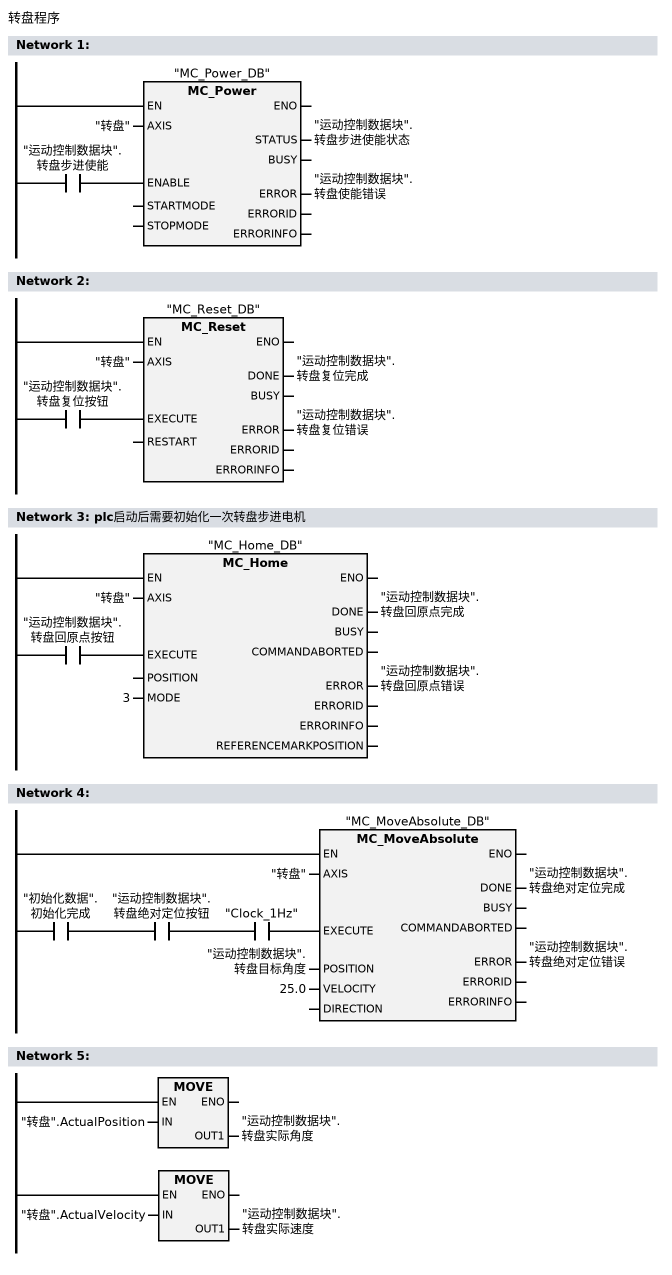
   "MC_Power_DB"(Axis := "转盘",   // MC_Power
                 Enable := "运动控制数据块".转盘步进使能,
                 Status => "运动控制数据块".转盘步进使能状态,
                 Error => "运动控制数据块".转盘使能错误);
END_REGION

REGION Network 2
   "MC_Reset_DB"(Axis := "转盘", Execute := "运动控制数据块".转盘复位按钮, Done => "运动控制数据块".转盘复位完成, Error => "运动控制数据块".转盘复位错误);   // MC_Reset
END_REGION

REGION Network 3: plc启动后需要初始化一次转盘步进电机
   "MC_Home_DB"(Axis := "转盘",   // MC_Home
                Execute := "运动控制数据块".转盘回原点按钮,
                Mode := 3,
                Done => "运动控制数据块".转盘回原点完成,
                Error => "运动控制数据块".转盘回原点错误);
END_REGION

REGION Network 4
   "MC_MoveAbsolute_DB"(Axis := "转盘",   // MC_MoveAbsolute
                        Execute := "初始化数据".初始化完成 AND "运动控制数据块".转盘绝对定位按钮 AND "Clock_1Hz",
                        Position := "运动控制数据块".转盘目标角度,
                        Velocity := 25.0,
                        Done => "运动控制数据块".转盘绝对定位完成,
                        Error => "运动控制数据块".转盘绝对定位错误);
END_REGION

REGION Network 5
   RUNG wire#powerrail
      Move(in := "转盘".ActualPosition, out1 => "运动控制数据块".转盘实际角度)
   END_RUNG
   RUNG wire#powerrail
      Move(in := "转盘".ActualVelocity, out1 => "运动控制数据块".转盘实际速度)
   END_RUNG
   // the same network as SCL:
   "运动控制数据块".转盘实际角度 := "转盘".ActualPosition;
   "运动控制数据块".转盘实际速度 := "转盘".ActualVelocity;
END_REGION
END_FUNCTION

FUNCTION "机械手程序" : Void   // FC8, LAD
{ S7_Optimized_Access := 'TRUE' }
VERSION : 0.1
// 极限位：左100，右-180
BEGIN

REGION Network 1: 轴使能
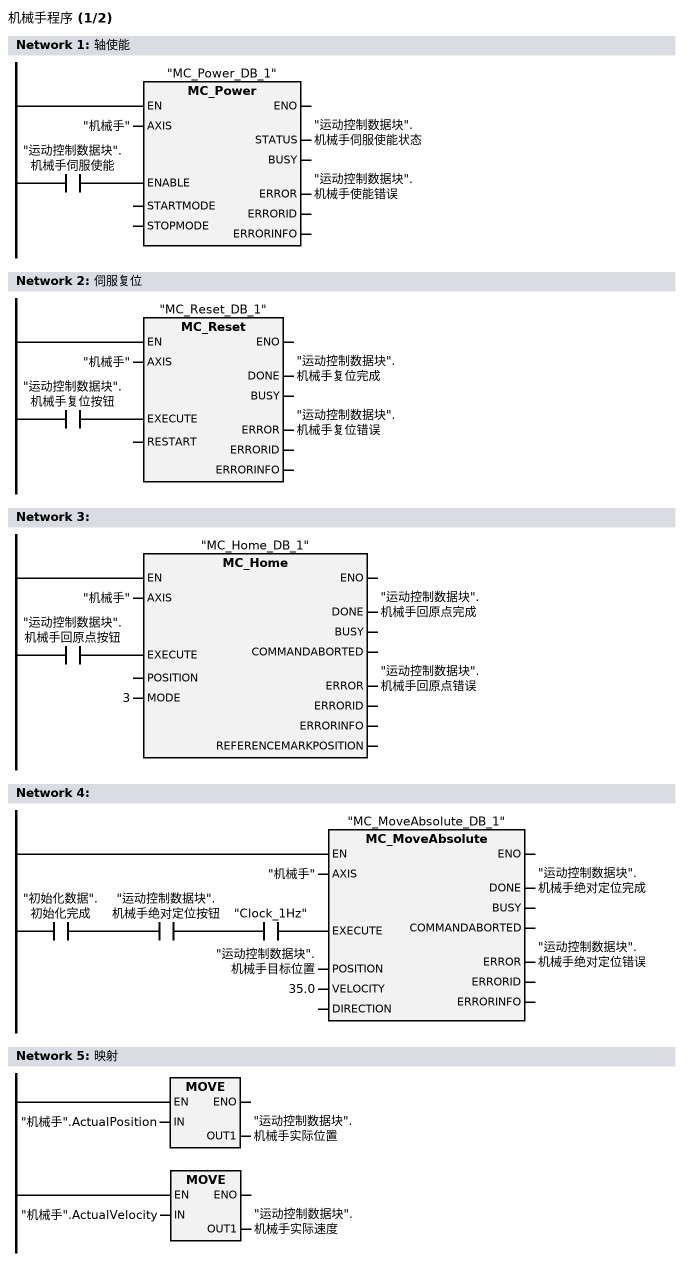
   "MC_Power_DB_1"(Axis := "机械手",   // MC_Power
                   Enable := "运动控制数据块".机械手伺服使能,
                   Status => "运动控制数据块".机械手伺服使能状态,
                   Error => "运动控制数据块".机械手使能错误);
END_REGION

REGION Network 2: 伺服复位
   "MC_Reset_DB_1"(Axis := "机械手",   // MC_Reset
                   Execute := "运动控制数据块".机械手复位按钮,
                   Done => "运动控制数据块".机械手复位完成,
                   Error => "运动控制数据块".机械手复位错误);
END_REGION

REGION Network 3
   "MC_Home_DB_1"(Axis := "机械手",   // MC_Home
                  Execute := "运动控制数据块".机械手回原点按钮,
                  Mode := 3,
                  Done => "运动控制数据块".机械手回原点完成,
                  Error => "运动控制数据块".机械手回原点错误);
END_REGION

REGION Network 4
   "MC_MoveAbsolute_DB_1"(Axis := "机械手",   // MC_MoveAbsolute
                          Execute := "初始化数据".初始化完成 AND "运动控制数据块".机械手绝对定位按钮 AND "Clock_1Hz",
                          Position := "运动控制数据块".机械手目标位置,
                          Velocity := 35.0,
                          Done => "运动控制数据块".机械手绝对定位完成,
                          Error => "运动控制数据块".机械手绝对定位错误);
END_REGION

REGION Network 5: 映射
   RUNG wire#powerrail
      Move(in := "机械手".ActualPosition, out1 => "运动控制数据块".机械手实际位置)
   END_RUNG
   RUNG wire#powerrail
      Move(in := "机械手".ActualVelocity, out1 => "运动控制数据块".机械手实际速度)
   END_RUNG
   // the same network as SCL:
   "运动控制数据块".机械手实际位置 := "机械手".ActualPosition;
   "运动控制数据块".机械手实际速度 := "机械手".ActualVelocity;
END_REGION

REGION Network 6
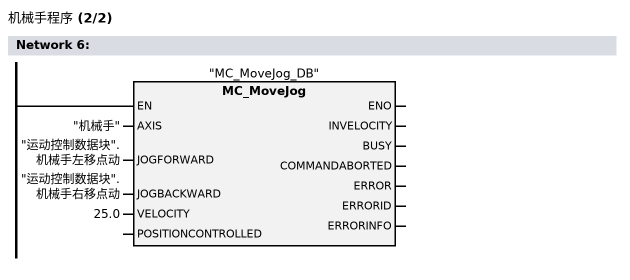
   "MC_MoveJog_DB"(Axis := "机械手",   // MC_MoveJog
                   JogForward := "运动控制数据块".机械手左移点动,
                   JogBackward := "运动控制数据块".机械手右移点动,
                   Velocity := 25.0);
END_REGION
END_FUNCTION

FUNCTION "[00]轴回零" : Void   // FC9, LAD
{ S7_Optimized_Access := 'TRUE' }
VERSION : 0.1
   VAR_TEMP   // added for the SCL form of the ladder/FBD networks
      _w1 : Bool;
   END_VAR
BEGIN

REGION Network 1
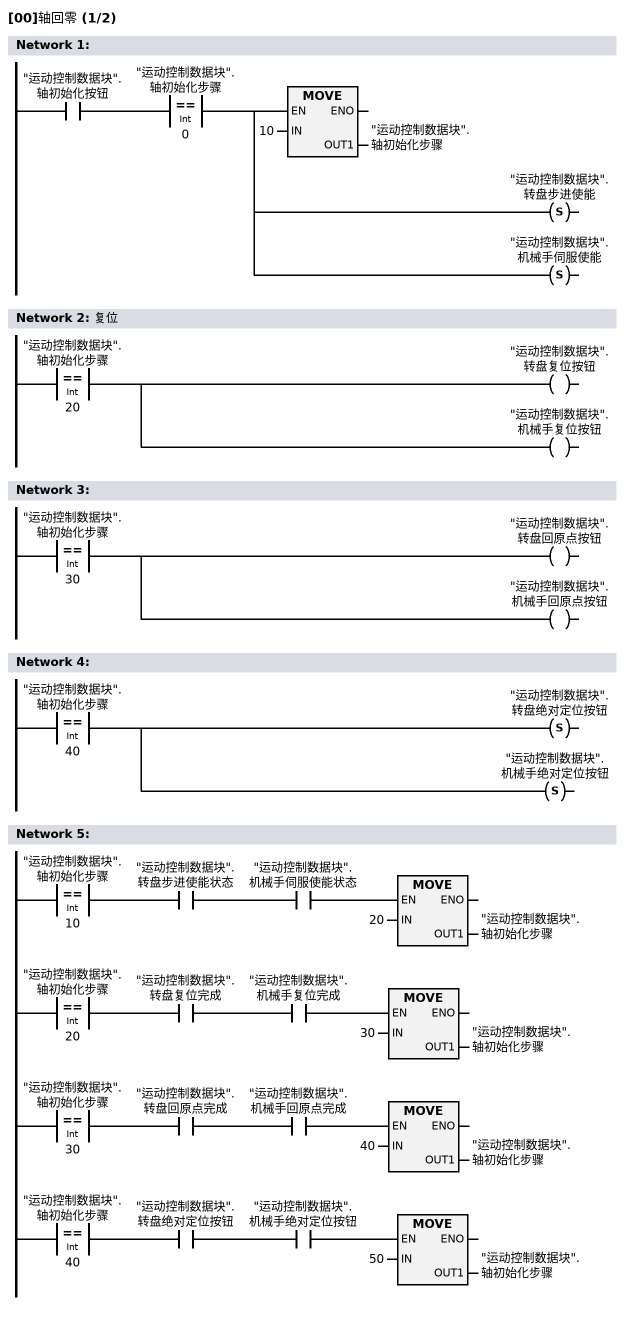
   RUNG wire#powerrail
      Contact( "运动控制数据块".轴初始化按钮 )
      { S7_Templates := "SrcType := Int" } EQ_Contact(in1 := "运动控制数据块".轴初始化步骤, in2 := 0)
      wire#w1
      Move(in := 10, out1 => "运动控制数据块".轴初始化步骤)
   END_RUNG
   RUNG wire#w1
      S_Coil( "运动控制数据块".转盘步进使能 )
   END_RUNG
   RUNG wire#w1
      S_Coil( "运动控制数据块".机械手伺服使能 )
   END_RUNG
   // the same network as SCL:
   #_w1 := "运动控制数据块".轴初始化按钮 AND ("运动控制数据块".轴初始化步骤 = 0);
   IF #_w1 THEN
       "运动控制数据块".轴初始化步骤 := 10;
       "运动控制数据块".转盘步进使能 := TRUE;
       "运动控制数据块".机械手伺服使能 := TRUE;
   END_IF;
END_REGION

REGION Network 2: 复位
   RUNG wire#powerrail
      { S7_Templates := "SrcType := Int" } EQ_Contact(in1 := "运动控制数据块".轴初始化步骤, in2 := 20)
      wire#w1
      Coil( "运动控制数据块".转盘复位按钮 )
   END_RUNG
   RUNG wire#w1
      Coil( "运动控制数据块".机械手复位按钮 )
   END_RUNG
   // the same network as SCL:
   "运动控制数据块".转盘复位按钮 := "运动控制数据块".轴初始化步骤 = 20;
   "运动控制数据块".机械手复位按钮 := "运动控制数据块".转盘复位按钮;
END_REGION

REGION Network 3
   RUNG wire#powerrail
      { S7_Templates := "SrcType := Int" } EQ_Contact(in1 := "运动控制数据块".轴初始化步骤, in2 := 30)
      wire#w1
      Coil( "运动控制数据块".转盘回原点按钮 )
   END_RUNG
   RUNG wire#w1
      Coil( "运动控制数据块".机械手回原点按钮 )
   END_RUNG
   // the same network as SCL:
   "运动控制数据块".转盘回原点按钮 := "运动控制数据块".轴初始化步骤 = 30;
   "运动控制数据块".机械手回原点按钮 := "运动控制数据块".转盘回原点按钮;
END_REGION

REGION Network 4
   RUNG wire#powerrail
      { S7_Templates := "SrcType := Int" } EQ_Contact(in1 := "运动控制数据块".轴初始化步骤, in2 := 40)
      wire#w1
      S_Coil( "运动控制数据块".转盘绝对定位按钮 )
   END_RUNG
   RUNG wire#w1
      S_Coil( "运动控制数据块".机械手绝对定位按钮 )
   END_RUNG
   // the same network as SCL:
   IF "运动控制数据块".轴初始化步骤 = 40 THEN
       "运动控制数据块".转盘绝对定位按钮 := TRUE;
       "运动控制数据块".机械手绝对定位按钮 := TRUE;
   END_IF;
END_REGION

REGION Network 5
   RUNG wire#powerrail
      { S7_Templates := "SrcType := Int" } EQ_Contact(in1 := "运动控制数据块".轴初始化步骤, in2 := 10)
      Contact( "运动控制数据块".转盘步进使能状态 )
      Contact( "运动控制数据块".机械手伺服使能状态 )
      Move(in := 20, out1 => "运动控制数据块".轴初始化步骤)
   END_RUNG
   RUNG wire#powerrail
      { S7_Templates := "SrcType := Int" } EQ_Contact(in1 := "运动控制数据块".轴初始化步骤, in2 := 20)
      Contact( "运动控制数据块".转盘复位完成 )
      Contact( "运动控制数据块".机械手复位完成 )
      Move(in := 30, out1 => "运动控制数据块".轴初始化步骤)
   END_RUNG
   RUNG wire#powerrail
      { S7_Templates := "SrcType := Int" } EQ_Contact(in1 := "运动控制数据块".轴初始化步骤, in2 := 30)
      Contact( "运动控制数据块".转盘回原点完成 )
      Contact( "运动控制数据块".机械手回原点完成 )
      Move(in := 40, out1 => "运动控制数据块".轴初始化步骤)
   END_RUNG
   RUNG wire#powerrail
      { S7_Templates := "SrcType := Int" } EQ_Contact(in1 := "运动控制数据块".轴初始化步骤, in2 := 40)
      Contact( "运动控制数据块".转盘绝对定位按钮 )
      Contact( "运动控制数据块".机械手绝对定位按钮 )
      Move(in := 50, out1 => "运动控制数据块".轴初始化步骤)
   END_RUNG
   // the same network as SCL:
   IF ("运动控制数据块".轴初始化步骤 = 10) AND "运动控制数据块".转盘步进使能状态 AND "运动控制数据块".机械手伺服使能状态 THEN
       "运动控制数据块".轴初始化步骤 := 20;
   END_IF;
   IF ("运动控制数据块".轴初始化步骤 = 20) AND "运动控制数据块".转盘复位完成 AND "运动控制数据块".机械手复位完成 THEN "运动控制数据块".轴初始化步骤 := 30; END_IF;
   IF ("运动控制数据块".轴初始化步骤 = 30) AND "运动控制数据块".转盘回原点完成 AND "运动控制数据块".机械手回原点完成 THEN
       "运动控制数据块".轴初始化步骤 := 40;
   END_IF;
   IF ("运动控制数据块".轴初始化步骤 = 40) AND "运动控制数据块".转盘绝对定位按钮 AND "运动控制数据块".机械手绝对定位按钮 THEN
       "运动控制数据块".轴初始化步骤 := 50;
   END_IF;
END_REGION

REGION Network 6: 轴初始化完成
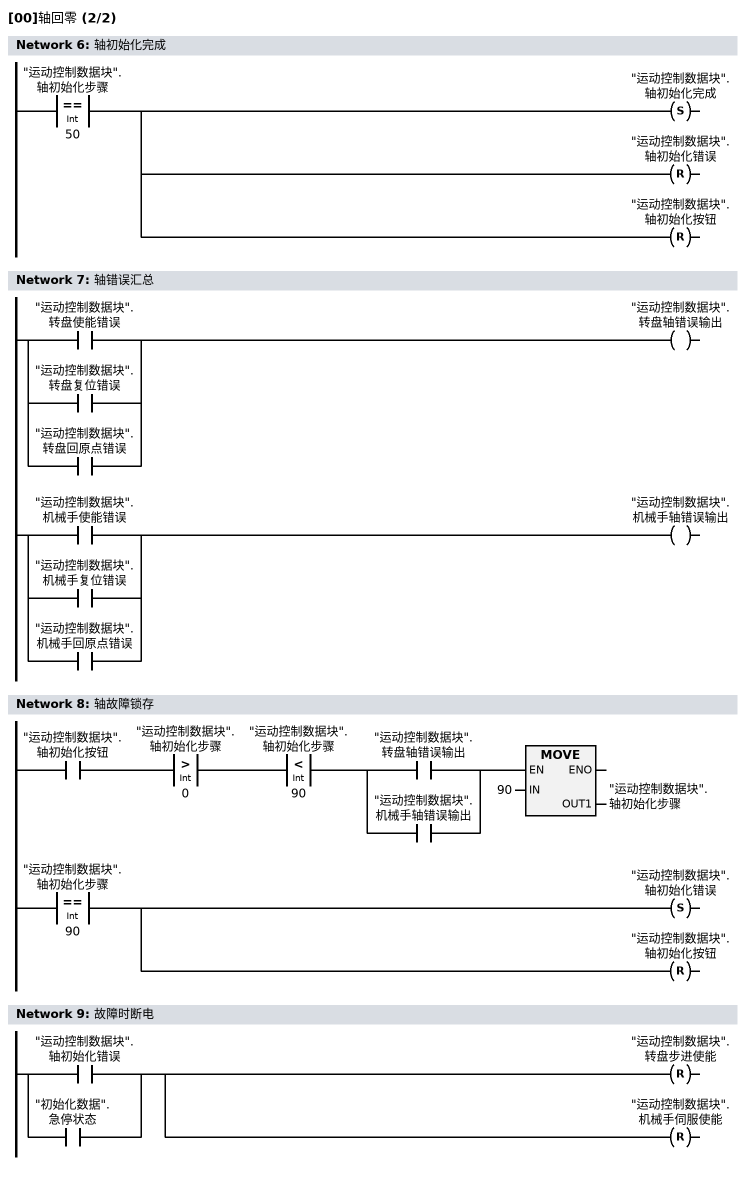
   RUNG wire#powerrail
      { S7_Templates := "SrcType := Int" } EQ_Contact(in1 := "运动控制数据块".轴初始化步骤, in2 := 50)
      wire#w1
      S_Coil( "运动控制数据块".轴初始化完成 )
   END_RUNG
   RUNG wire#w1
      R_Coil( "运动控制数据块".轴初始化错误 )
   END_RUNG
   RUNG wire#w1
      R_Coil( "运动控制数据块".轴初始化按钮 )
   END_RUNG
   // the same network as SCL:
   IF "运动控制数据块".轴初始化步骤 = 50 THEN
       "运动控制数据块".轴初始化完成 := TRUE;
       "运动控制数据块".轴初始化错误 := FALSE;
       "运动控制数据块".轴初始化按钮 := FALSE;
   END_IF;
END_REGION

REGION Network 7: 轴错误汇总
   RUNG wire#powerrail
      Contact( "运动控制数据块".转盘使能错误 )
      wire#w1
      Coil( "运动控制数据块".转盘轴错误输出 )
   END_RUNG
   RUNG wire#powerrail
      Contact( "运动控制数据块".转盘复位错误 )
   END_RUNG wire#w1
   RUNG wire#powerrail
      Contact( "运动控制数据块".转盘回原点错误 )
   END_RUNG wire#w1
   RUNG wire#powerrail
      Contact( "运动控制数据块".机械手使能错误 )
      wire#w2
      Coil( "运动控制数据块".机械手轴错误输出 )
   END_RUNG
   RUNG wire#powerrail
      Contact( "运动控制数据块".机械手复位错误 )
   END_RUNG wire#w2
   RUNG wire#powerrail
      Contact( "运动控制数据块".机械手回原点错误 )
   END_RUNG wire#w2
   // the same network as SCL:
   "运动控制数据块".转盘轴错误输出 := "运动控制数据块".转盘使能错误 OR "运动控制数据块".转盘复位错误 OR "运动控制数据块".转盘回原点错误;
   "运动控制数据块".机械手轴错误输出 := "运动控制数据块".机械手使能错误 OR "运动控制数据块".机械手复位错误 OR "运动控制数据块".机械手回原点错误;
END_REGION

REGION Network 8: 轴故障锁存
   RUNG wire#powerrail
      Contact( "运动控制数据块".轴初始化按钮 )
      { S7_Templates := "SrcType := Int" } GT_Contact(in1 := "运动控制数据块".轴初始化步骤, in2 := 0)
      { S7_Templates := "SrcType := Int" } LT_Contact(in1 := "运动控制数据块".轴初始化步骤, in2 := 90)
      wire#w1
      Contact( "运动控制数据块".转盘轴错误输出 )
      wire#w2
      Move(in := 90, out1 => "运动控制数据块".轴初始化步骤)
   END_RUNG
   RUNG wire#w1
      Contact( "运动控制数据块".机械手轴错误输出 )
   END_RUNG wire#w2
   RUNG wire#powerrail
      { S7_Templates := "SrcType := Int" } EQ_Contact(in1 := "运动控制数据块".轴初始化步骤, in2 := 90)
      wire#w3
      S_Coil( "运动控制数据块".轴初始化错误 )
   END_RUNG
   RUNG wire#w3
      R_Coil( "运动控制数据块".轴初始化按钮 )
   END_RUNG
   // the same network as SCL:
   IF "运动控制数据块".轴初始化按钮 AND ("运动控制数据块".轴初始化步骤 > 0) AND ("运动控制数据块".轴初始化步骤 < 90) AND ("运动控制数据块".转盘轴错误输出 OR "运动控制数据块".机械手轴错误输出) THEN
       "运动控制数据块".轴初始化步骤 := 90;
   END_IF;
   IF "运动控制数据块".轴初始化步骤 = 90 THEN
       "运动控制数据块".轴初始化错误 := TRUE;
       "运动控制数据块".轴初始化按钮 := FALSE;
   END_IF;
END_REGION

REGION Network 9: 故障时断电
   RUNG wire#powerrail
      Contact( "运动控制数据块".轴初始化错误 )
      wire#w1
      R_Coil( "运动控制数据块".转盘步进使能 )
   END_RUNG
   RUNG wire#powerrail
      Contact( "初始化数据".急停状态 )
   END_RUNG wire#w1
   RUNG wire#w1
      R_Coil( "运动控制数据块".机械手伺服使能 )
   END_RUNG
   // the same network as SCL:
   IF "运动控制数据块".轴初始化错误 OR "初始化数据".急停状态 THEN
       "运动控制数据块".转盘步进使能 := FALSE;
       "运动控制数据块".机械手伺服使能 := FALSE;
   END_IF;
END_REGION
END_FUNCTION

// folder: 通讯数据

FUNCTION "产线通讯" : Void   // FC16, LAD
{ S7_Optimized_Access := 'TRUE' }
VERSION : 0.1
BEGIN

REGION Network 1: 心跳
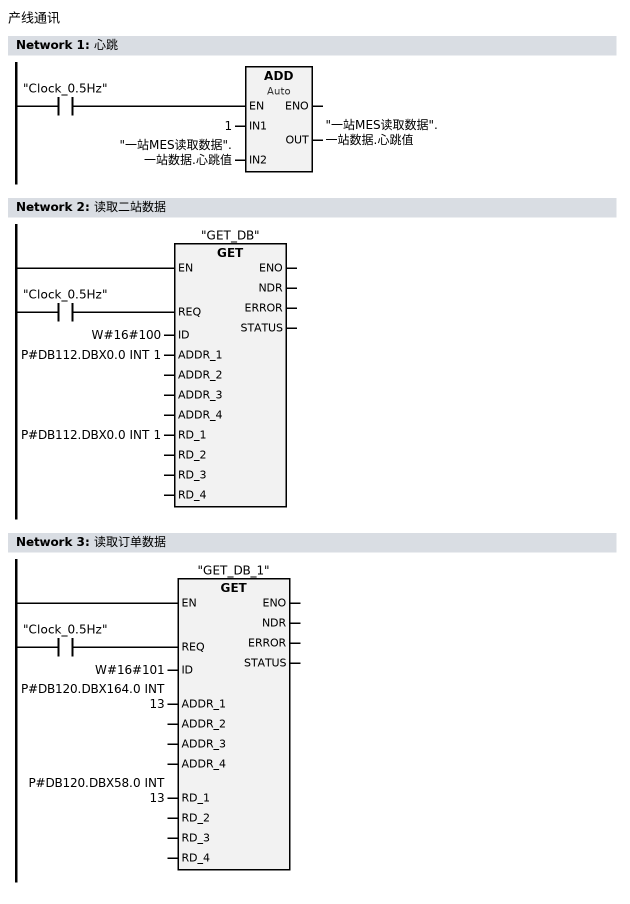
   RUNG wire#powerrail
      Contact( "Clock_0.5Hz" )
      Add(in1 := 1, in2 := "一站MES读取数据".一站数据.心跳值, out => "一站MES读取数据".一站数据.心跳值)
   END_RUNG
   // the same network as SCL:
   IF "Clock_0.5Hz" THEN "一站MES读取数据".一站数据.心跳值 := 1 + "一站MES读取数据".一站数据.心跳值; END_IF;
END_REGION

REGION Network 2: 读取二站数据
   "GET_DB"(REQ := "Clock_0.5Hz", ID := W#16#100, ADDR_1 := P#DB112.DBX0.0 INT 1, RD_1 := P#DB112.DBX0.0 INT 1);   // GET
END_REGION

REGION Network 3: 读取订单数据
   "GET_DB_1"(REQ := "Clock_0.5Hz",   // GET
              ID := W#16#101,
              ADDR_1 := P#DB120.DBX164.0 INT 13,
              RD_1 := P#DB120.DBX58.0 INT 13);
END_REGION
END_FUNCTION

FUNCTION "MES数据映射" : Void   // FC18, LAD
{ S7_Optimized_Access := 'TRUE' }
VERSION : 0.1
BEGIN

REGION Network 1: 运行模式
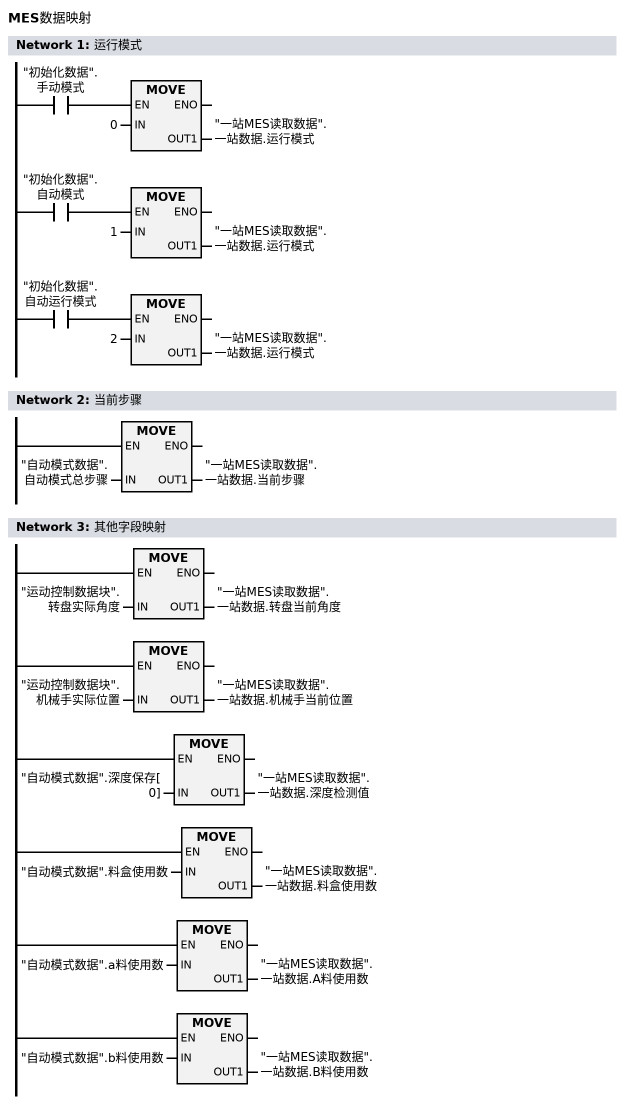
   RUNG wire#powerrail
      Contact( "初始化数据".手动模式 )
      Move(in := 0, out1 => "一站MES读取数据".一站数据.运行模式)
   END_RUNG
   RUNG wire#powerrail
      Contact( "初始化数据".自动模式 )
      Move(in := 1, out1 => "一站MES读取数据".一站数据.运行模式)
   END_RUNG
   RUNG wire#powerrail
      Contact( "初始化数据".自动运行模式 )
      Move(in := 2, out1 => "一站MES读取数据".一站数据.运行模式)
   END_RUNG
   // the same network as SCL:
   IF "初始化数据".手动模式 THEN "一站MES读取数据".一站数据.运行模式 := 0; END_IF;
   IF "初始化数据".自动模式 THEN "一站MES读取数据".一站数据.运行模式 := 1; END_IF;
   IF "初始化数据".自动运行模式 THEN "一站MES读取数据".一站数据.运行模式 := 2; END_IF;
END_REGION

REGION Network 2: 当前步骤
   RUNG wire#powerrail
      Move(in := "自动模式数据".自动模式总步骤, out1 => "一站MES读取数据".一站数据.当前步骤)
   END_RUNG
   // the same network as SCL:
   "一站MES读取数据".一站数据.当前步骤 := "自动模式数据".自动模式总步骤;
END_REGION

REGION Network 3: 其他字段映射
   RUNG wire#powerrail
      Move(in := "运动控制数据块".转盘实际角度, out1 => "一站MES读取数据".一站数据.转盘当前角度)
   END_RUNG
   RUNG wire#powerrail
      Move(in := "运动控制数据块".机械手实际位置, out1 => "一站MES读取数据".一站数据.机械手当前位置)
   END_RUNG
   RUNG wire#powerrail
      Move(in := "自动模式数据".深度保存[0], out1 => "一站MES读取数据".一站数据.深度检测值)
   END_RUNG
   RUNG wire#powerrail
      Move(in := "自动模式数据".料盒使用数, out1 => "一站MES读取数据".一站数据.料盒使用数)
   END_RUNG
   RUNG wire#powerrail
      Move(in := "自动模式数据".a料使用数, out1 => "一站MES读取数据".一站数据.A料使用数)
   END_RUNG
   RUNG wire#powerrail
      Move(in := "自动模式数据".b料使用数, out1 => "一站MES读取数据".一站数据.B料使用数)
   END_RUNG
   // the same network as SCL:
   "一站MES读取数据".一站数据.转盘当前角度 := "运动控制数据块".转盘实际角度;
   "一站MES读取数据".一站数据.机械手当前位置 := "运动控制数据块".机械手实际位置;
   "一站MES读取数据".一站数据.深度检测值 := "自动模式数据".深度保存[0];
   "一站MES读取数据".一站数据.料盒使用数 := "自动模式数据".料盒使用数;
   "一站MES读取数据".一站数据.A料使用数 := "自动模式数据".a料使用数;
   "一站MES读取数据".一站数据.B料使用数 := "自动模式数据".b料使用数;
END_REGION
END_FUNCTION

FUNCTION "扫码器通信" : Void   // FC19, LAD
{ S7_Optimized_Access := 'TRUE' }
VERSION : 0.1
BEGIN

REGION Network 1
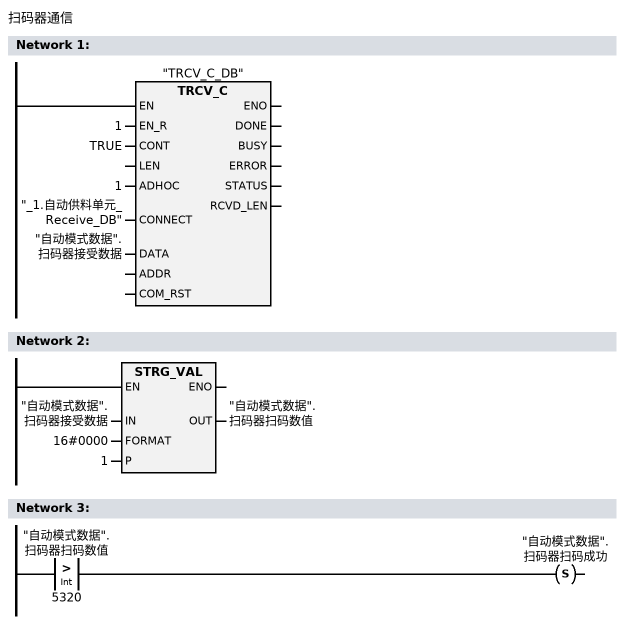
   "TRCV_C_DB"(EN_R := 1, CONT := TRUE, ADHOC := 1, CONNECT := "_1.自动供料单元_Receive_DB", DATA := "自动模式数据".扫码器接受数据);   // TRCV_C
END_REGION

REGION Network 2
   STRG_VAL(IN := "自动模式数据".扫码器接受数据, FORMAT := 16#0000, P := 1, OUT => "自动模式数据".扫码器扫码数值);
END_REGION

REGION Network 3
   RUNG wire#powerrail
      { S7_Templates := "SrcType := Int" } GT_Contact(in1 := "自动模式数据".扫码器扫码数值, in2 := 5320)
      S_Coil( "自动模式数据".扫码器扫码成功 )
   END_RUNG
   // the same network as SCL:
   IF "自动模式数据".扫码器扫码数值 > 5320 THEN "自动模式数据".扫码器扫码成功 := TRUE; END_IF;
END_REGION
END_FUNCTION

FUNCTION "虚实联动映射" : Void   // FC20, LAD
{ S7_Optimized_Access := 'TRUE' }
VERSION : 0.1
BEGIN

REGION Network 1
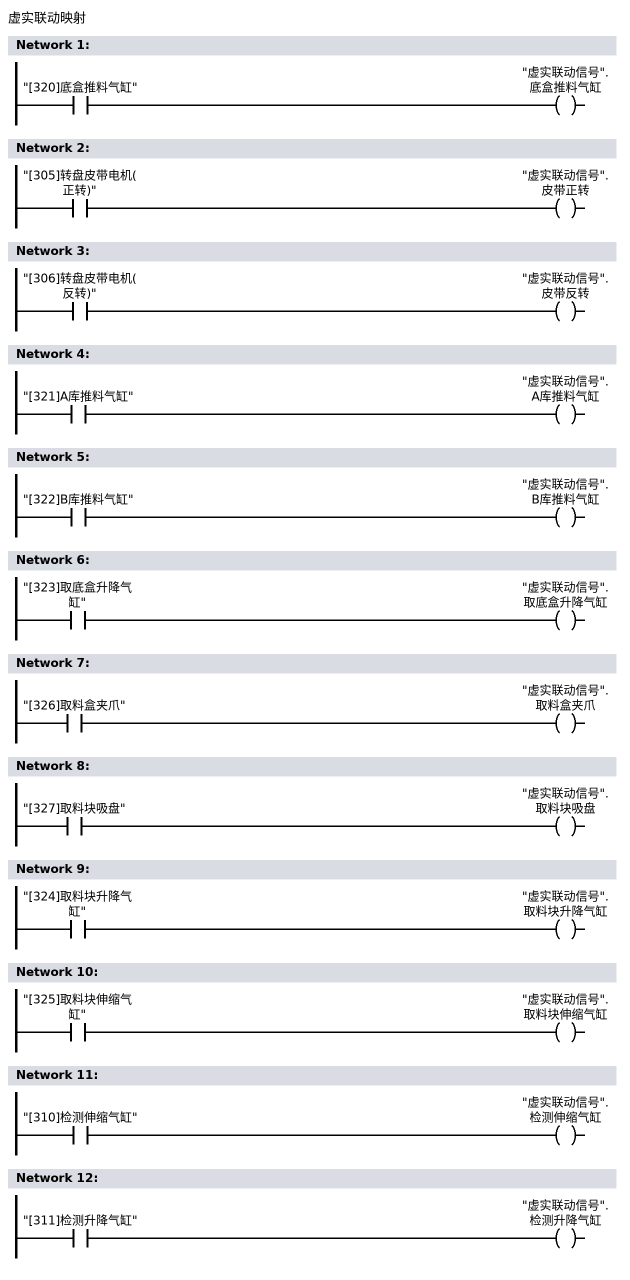
   RUNG wire#powerrail
      Contact( "[320]底盒推料气缸" )
      Coil( "虚实联动信号".底盒推料气缸 )
   END_RUNG
   // the same network as SCL:
   "虚实联动信号".底盒推料气缸 := "[320]底盒推料气缸";
END_REGION

REGION Network 2
   RUNG wire#powerrail
      Contact( "[305]转盘皮带电机(正转)" )
      Coil( "虚实联动信号".皮带正转 )
   END_RUNG
   // the same network as SCL:
   "虚实联动信号".皮带正转 := "[305]转盘皮带电机(正转)";
END_REGION

REGION Network 3
   RUNG wire#powerrail
      Contact( "[306]转盘皮带电机(反转)" )
      Coil( "虚实联动信号".皮带反转 )
   END_RUNG
   // the same network as SCL:
   "虚实联动信号".皮带反转 := "[306]转盘皮带电机(反转)";
END_REGION

REGION Network 4
   RUNG wire#powerrail
      Contact( "[321]A库推料气缸" )
      Coil( "虚实联动信号".A库推料气缸 )
   END_RUNG
   // the same network as SCL:
   "虚实联动信号".A库推料气缸 := "[321]A库推料气缸";
END_REGION

REGION Network 5
   RUNG wire#powerrail
      Contact( "[322]B库推料气缸" )
      Coil( "虚实联动信号".B库推料气缸 )
   END_RUNG
   // the same network as SCL:
   "虚实联动信号".B库推料气缸 := "[322]B库推料气缸";
END_REGION

REGION Network 6
   RUNG wire#powerrail
      Contact( "[323]取底盒升降气缸" )
      Coil( "虚实联动信号".取底盒升降气缸 )
   END_RUNG
   // the same network as SCL:
   "虚实联动信号".取底盒升降气缸 := "[323]取底盒升降气缸";
END_REGION

REGION Network 7
   RUNG wire#powerrail
      Contact( "[326]取料盒夹爪" )
      Coil( "虚实联动信号".取料盒夹爪 )
   END_RUNG
   // the same network as SCL:
   "虚实联动信号".取料盒夹爪 := "[326]取料盒夹爪";
END_REGION

REGION Network 8
   RUNG wire#powerrail
      Contact( "[327]取料块吸盘" )
      Coil( "虚实联动信号".取料块吸盘 )
   END_RUNG
   // the same network as SCL:
   "虚实联动信号".取料块吸盘 := "[327]取料块吸盘";
END_REGION

REGION Network 9
   RUNG wire#powerrail
      Contact( "[324]取料块升降气缸" )
      Coil( "虚实联动信号".取料块升降气缸 )
   END_RUNG
   // the same network as SCL:
   "虚实联动信号".取料块升降气缸 := "[324]取料块升降气缸";
END_REGION

REGION Network 10
   RUNG wire#powerrail
      Contact( "[325]取料块伸缩气缸" )
      Coil( "虚实联动信号".取料块伸缩气缸 )
   END_RUNG
   // the same network as SCL:
   "虚实联动信号".取料块伸缩气缸 := "[325]取料块伸缩气缸";
END_REGION

REGION Network 11
   RUNG wire#powerrail
      Contact( "[310]检测伸缩气缸" )
      Coil( "虚实联动信号".检测伸缩气缸 )
   END_RUNG
   // the same network as SCL:
   "虚实联动信号".检测伸缩气缸 := "[310]检测伸缩气缸";
END_REGION

REGION Network 12
   RUNG wire#powerrail
      Contact( "[311]检测升降气缸" )
      Coil( "虚实联动信号".检测升降气缸 )
   END_RUNG
   // the same network as SCL:
   "虚实联动信号".检测升降气缸 := "[311]检测升降气缸";
END_REGION
END_FUNCTION

// ===== PLC "2.智能分拣单元"  CPU 1214C DC/DC/DC =====

VAR_GLOBAL   // PLC tag table "默认变量表"
   "System_Byte" AT %MB501 : Byte;
   "FirstScan" AT %M501.0 : Bool;
   "DiagStatusUpdate" AT %M501.1 : Bool;
   "AlwaysTRUE" AT %M501.2 : Bool;
   "AlwaysFALSE" AT %M501.3 : Bool;
   "Clock_Byte" AT %MB500 : Byte;
   "Clock_10Hz" AT %M500.0 : Bool;
   "Clock_5Hz" AT %M500.1 : Bool;
   "Clock_2.5Hz" AT %M500.2 : Bool;
   "Clock_2Hz" AT %M500.3 : Bool;
   "Clock_1.25Hz" AT %M500.4 : Bool;
   "Clock_1Hz" AT %M500.5 : Bool;
   "Clock_0.625Hz" AT %M500.6 : Bool;
   "Clock_0.5Hz" AT %M500.7 : Bool;
   "Tag_1" AT %M5.1 : Bool;
   "注释按钮" AT %M100.0 : Bool;
END_VAR

VAR_GLOBAL   // PLC tag table "第二站变量表"
   "[100]启动" AT %I0.0 : Bool;
   "[101]停止" AT %I0.1 : Bool;
   "[102]复位" AT %I0.2 : Bool;
   "[103]急停" AT %I0.3 : Bool;
   "[104]手自动" AT %I0.4 : Bool;
   "[105]8mm钢球检测" AT %I0.5 : Bool;
   "[107]备用" AT %I0.7 : Bool;
   "[110]备用" AT %I1.0 : Bool;
   "[111]备用" AT %I1.1 : Bool;
   "[112]备用" AT %I1.2 : Bool;
   "[113]备用" AT %I1.3 : Bool;
   "[114]备用" AT %I1.4 : Bool;
   "[120]8mm挡停缩回" AT %I2.0 : Bool;
   "[121]8mm挡停伸出" AT %I2.1 : Bool;
   "[122]8mm料盒到达" AT %I2.2 : Bool;
   "[123]8mm推料缩回" AT %I2.3 : Bool;
   "传输伺服_Drive_OUT" AT %Q64.0 : "PD_TEL3_OUT";
   "[300]8mm分拣步进_脉冲" AT %Q0.0 : Bool;
   "[301]10mm分拣步进_脉冲" AT %Q0.1 : Bool;
   "[302]8mm分拣步进_方向" AT %Q0.2 : Bool;
   "[303]10mm分拣步进_方向" AT %Q0.3 : Bool;
   "[320]8mm挡停气缸" AT %Q2.0 : Bool;
   "[321]8mm推料气缸" AT %Q2.1 : Bool;   // 0为伸出，1为缩回，伸出时料仓检测有效
   "[322]10mm挡停气缸" AT %Q2.2 : Bool;
   "[323]10mm推料气缸" AT %Q2.3 : Bool;
   "[324]备用" AT %Q2.4 : Bool;
   "[325]备用" AT %Q2.5 : Bool;
   "[326]备用" AT %Q2.6 : Bool;
   "[327]备用" AT %Q2.7 : Bool;
   "[124]8mm柱状料仓有无" AT %I2.4 : Bool;
   "[125]10mm挡停缩回" AT %I2.5 : Bool;
   "[115]备用" AT %I1.5 : Bool;
   "[106]10mm钢球检测" AT %I0.6 : Bool;
   "[304]黄色指示灯" AT %Q0.4 : Bool;
   "[305]绿色指示灯" AT %Q0.5 : Bool;
   "[306]红色指示灯" AT %Q0.6 : Bool;
   "[307]声光报警" AT %Q0.7 : Bool;
   "[310]备用" AT %Q1.0 : Bool;
   "[311]备用" AT %Q1.1 : Bool;
   "[156]光栅开关" AT %I5.6 : Bool;
   "[164]深度检测" AT %IW64 : Word;
   "传输伺服_Drive_IN(1)" AT %I68.0 : "PD_TEL3_IN";
   "[126]10mm挡停伸出" AT %I2.6 : Bool;
   "[127]10mm料盒到达" AT %I2.7 : Bool;
   "[130]10mm推料缩回" AT %I3.0 : Bool;
   "[131]10mm柱状料仓有无" AT %I3.1 : Bool;
END_VAR

DATA_BLOCK "初始化数据"   // DB19
{ S7_Optimized_Access := 'FALSE' }
VERSION : 0.1
   VAR
      初始化步骤 : Int;
      初始化完成 : Bool;
      初始化中 : Bool;
      初始化故障 : Bool;
      急停状态 : Bool;
      复位完成 : Bool;
      手动模式 : Bool;
      自动模式 : Bool;
      自动运行模式 : Bool;
      黄灯_内部 : Bool;
      红灯_内部 : Bool;
      绿灯_内部 : Bool;
      安全光栅被挡 : Bool;
      报警等级 : Int;
      报警确认按钮 : Bool;
      "8mm挡停气缸报警" : Bool;
      "10mm挡停气缸报警" : Bool;
      报警总输出 : Bool;
      报警状态确认 : Bool;
   END_VAR
BEGIN
END_DATA_BLOCK

DATA_BLOCK "状态控制数据"   // DB28
{ S7_Optimized_Access := 'FALSE' }
VERSION : 0.1
   VAR
      在线状态 : Bool;
      空闲状态 : Bool;
      忙碌状态 : Bool;
      故障状态 : Bool;
   END_VAR
BEGIN
END_DATA_BLOCK

DATA_BLOCK "二站MES读取数据"   // DB120
{ S7_Optimized_Access := 'FALSE' }
VERSION : 0.1
   VAR
      二站数据 : Struct
         在线状态 : Int;
         运行模式 : Int;   // 0 手动 / 1 自动待机 / 2 自动运行
         忙碌状态 : Int;   // 0 空闲 / 1 忙碌
         故障状态 : Int;   // 0 = 无故障
         当前订单ID : Int;   // 当前处理的订单
         当前步骤 : Real;
         心跳值 : Int;
         二站完成 : Bool;
         保留 : Bool;
         保留_1 : Bool;
         保留_2 : Bool;
         保留_3 : Bool;
         保留_4 : Bool;
         保留_5 : Bool;
         保留_6 : Bool;
         二站扫码数据 : Int;
         "8mm已灌注数量" : Int;
         "10mm已灌注数量" : Int;
         "8mml料仓钢珠有无" : Bool;   // 1有0无
         "10mm料仓钢珠有无" : Bool;   // 1有0无
         二站保留数据 : Array[0..9] of Int;
      END_STRUCT;
      订单数据 : Struct
         订单id : Int;
         ab物料 : Int;   // 1A，2B，3不需要
         小钢珠数量 : Int;
         大钢珠数量 : Int;
         存储仓位 : Int;
         当前订单完成 : Bool;
         开始信号 : Int;
         复位信号 : Int;
         订单保留数据 : Array[0..4] of Int;
      END_STRUCT;
   END_VAR
BEGIN
END_DATA_BLOCK

// folder: System blocks/Program resources

DATA_BLOCK "IEC_Timer_0_DB_16"   // DB3
{ S7_Optimized_Access := 'TRUE' }
AUTHOR : Simatic
FAMILY : IEC
NAME : IEC_TMR
VERSION : 1.0
// stored: InstanceOfName IEC_TIMER
"IEC_TIMER"
BEGIN
END_DATA_BLOCK

DATA_BLOCK "IEC_Timer_0_DB"   // DB4
{ S7_Optimized_Access := 'TRUE' }
AUTHOR : Simatic
FAMILY : IEC
NAME : IEC_TMR
VERSION : 1.0
// stored: InstanceOfName IEC_TIMER
"IEC_TIMER"
BEGIN
END_DATA_BLOCK

DATA_BLOCK "IEC_Timer_0_DB_1"   // DB5
{ S7_Optimized_Access := 'TRUE' }
AUTHOR : Simatic
FAMILY : IEC
NAME : IEC_TMR
VERSION : 1.0
// stored: InstanceOfName IEC_TIMER
"IEC_TIMER"
BEGIN
END_DATA_BLOCK

DATA_BLOCK "IEC_Timer_0_DB_2"   // DB7
{ S7_Optimized_Access := 'TRUE' }
AUTHOR : Simatic
FAMILY : IEC
NAME : IEC_TMR
VERSION : 1.0
// stored: InstanceOfName IEC_TIMER
"IEC_TIMER"
BEGIN
END_DATA_BLOCK

DATA_BLOCK "IEC_Timer_0_DB_3"   // DB8
{ S7_Optimized_Access := 'TRUE' }
AUTHOR : Simatic
FAMILY : IEC
NAME : IEC_TMR
VERSION : 1.0
// stored: InstanceOfName IEC_TIMER
"IEC_TIMER"
BEGIN
END_DATA_BLOCK

DATA_BLOCK "IEC_Timer_0_DB_4"   // DB9
{ S7_Optimized_Access := 'TRUE' }
AUTHOR : Simatic
FAMILY : IEC
NAME : IEC_TMR
VERSION : 1.0
// stored: InstanceOfName IEC_TIMER
"IEC_TIMER"
BEGIN
END_DATA_BLOCK

DATA_BLOCK "IEC_Timer_0_DB_5"   // DB10
{ S7_Optimized_Access := 'TRUE' }
AUTHOR : Simatic
FAMILY : IEC
NAME : IEC_TMR
VERSION : 1.0
// stored: InstanceOfName IEC_TIMER
"IEC_TIMER"
BEGIN
END_DATA_BLOCK

DATA_BLOCK "IEC_Timer_0_DB_6"   // DB11
{ S7_Optimized_Access := 'TRUE' }
AUTHOR : Simatic
FAMILY : IEC
NAME : IEC_TMR
VERSION : 1.0
// stored: InstanceOfName IEC_TIMER
"IEC_TIMER"
BEGIN
END_DATA_BLOCK

DATA_BLOCK "IEC_Timer_0_DB_7"   // DB12
{ S7_Optimized_Access := 'TRUE' }
AUTHOR : Simatic
FAMILY : IEC
NAME : IEC_TMR
VERSION : 1.0
// stored: InstanceOfName IEC_TIMER
"IEC_TIMER"
BEGIN
END_DATA_BLOCK

DATA_BLOCK "IEC_Timer_0_DB_8"   // DB13
{ S7_Optimized_Access := 'TRUE' }
AUTHOR : Simatic
FAMILY : IEC
NAME : IEC_TMR
VERSION : 1.0
// stored: InstanceOfName IEC_TIMER
"IEC_TIMER"
BEGIN
END_DATA_BLOCK

DATA_BLOCK "IEC_Timer_0_DB_9"   // DB14
{ S7_Optimized_Access := 'TRUE' }
AUTHOR : Simatic
FAMILY : IEC
NAME : IEC_TMR
VERSION : 1.0
// stored: InstanceOfName IEC_TIMER
"IEC_TIMER"
BEGIN
END_DATA_BLOCK

DATA_BLOCK "_2.智能分拣单元_Receive_DB"   // DB16
{ S7_Optimized_Access := 'TRUE' }
AUTHOR : SIMATIC
FAMILY : MC7Plus
NAME : TC_IP_v4
VERSION : 1.0
// stored: InstanceOfName TCON_IP_v4
"TCON_IP_v4"
BEGIN
   ID := 110;
   InterfaceId := 64;
   LocalPort := 8899;
   RemotePort := 8899;
   RemoteAddress.ADDR[1] := 192;
   RemoteAddress.ADDR[2] := 168;
   RemoteAddress.ADDR[3] := 40;
   RemoteAddress.ADDR[4] := 101;
END_DATA_BLOCK

DATA_BLOCK "IEC_Timer_0_DB_10"   // DB17
{ S7_Optimized_Access := 'TRUE' }
AUTHOR : Simatic
FAMILY : IEC
NAME : IEC_TMR
VERSION : 1.0
// stored: InstanceOfName IEC_TIMER
"IEC_TIMER"
BEGIN
END_DATA_BLOCK

DATA_BLOCK "IEC_Timer_0_DB_11"   // DB18
{ S7_Optimized_Access := 'TRUE' }
AUTHOR : Simatic
FAMILY : IEC
NAME : IEC_TMR
VERSION : 1.0
// stored: InstanceOfName IEC_TIMER
"IEC_TIMER"
BEGIN
END_DATA_BLOCK

DATA_BLOCK "IEC_Timer_0_DB_12"   // DB20
{ S7_Optimized_Access := 'TRUE' }
AUTHOR : Simatic
FAMILY : IEC
NAME : IEC_TMR
VERSION : 1.0
// stored: InstanceOfName IEC_TIMER
"IEC_TIMER"
BEGIN
END_DATA_BLOCK

DATA_BLOCK "IEC_Timer_0_DB_13"   // DB21
{ S7_Optimized_Access := 'TRUE' }
AUTHOR : Simatic
FAMILY : IEC
NAME : IEC_TMR
VERSION : 1.0
// stored: InstanceOfName IEC_TIMER
"IEC_TIMER"
BEGIN
END_DATA_BLOCK

DATA_BLOCK "IEC_Timer_0_DB_14"   // DB22
{ S7_Optimized_Access := 'TRUE' }
AUTHOR : Simatic
FAMILY : IEC
NAME : IEC_TMR
VERSION : 1.0
// stored: InstanceOfName IEC_TIMER
"IEC_TIMER"
BEGIN
END_DATA_BLOCK

DATA_BLOCK "IEC_Timer_0_DB_15"   // DB23
{ S7_Optimized_Access := 'TRUE' }
AUTHOR : Simatic
FAMILY : IEC
NAME : IEC_TMR
VERSION : 1.0
// stored: InstanceOfName IEC_TIMER
"IEC_TIMER"
BEGIN
END_DATA_BLOCK

DATA_BLOCK "IEC_Timer_0_DB_19"   // DB25
{ S7_Optimized_Access := 'TRUE' }
AUTHOR : Simatic
FAMILY : IEC
NAME : IEC_TMR
VERSION : 1.0
// stored: InstanceOfName IEC_TIMER
"IEC_TIMER"
BEGIN
END_DATA_BLOCK

DATA_BLOCK "IEC_Timer_0_DB_17"   // DB26
{ S7_Optimized_Access := 'TRUE' }
AUTHOR : Simatic
FAMILY : IEC
NAME : IEC_TMR
VERSION : 1.0
// stored: InstanceOfName IEC_TIMER
"IEC_TIMER"
BEGIN
END_DATA_BLOCK

DATA_BLOCK "IEC_Timer_0_DB_18"   // DB27
{ S7_Optimized_Access := 'TRUE' }
AUTHOR : Simatic
FAMILY : IEC
NAME : IEC_TMR
VERSION : 1.0
// stored: InstanceOfName IEC_TIMER
"IEC_TIMER"
BEGIN
END_DATA_BLOCK

// folder: 手动模式

DATA_BLOCK "手动模式数据"   // DB1
{ S7_Optimized_Access := 'FALSE' }
VERSION : 0.1
   VAR
      手动灌注总步骤 : Real;
      "8mm灌料步骤" : Real;
      "8mm现有钢珠" : Int;
      "8mm目标数量" : Int;
      "8mm灌注完成" : Bool;
      "10mm灌料步骤" : Real;
      "10mm现有钢珠" : Int;
      "10mm目标数量" : Int;
      "10mm灌注完成" : Bool;
   END_VAR
BEGIN
END_DATA_BLOCK

// folder: 自动模式

DATA_BLOCK "自动模式数据"   // DB6
{ S7_Optimized_Access := 'FALSE' }
VERSION : 0.1
   VAR
      自动灌注总步骤 : Real;
      "8mm灌料步骤" : Real;
      "8mm现有钢珠" : Int;
      "8mm下单数量" : Int;
      "8mm灌注完成" : Bool;
      "10mm灌料步骤" : Real;
      "10mm现有钢珠" : Int;
      "10mm下单数量" : Int;
      "10mm灌注完成" : Bool;
      检测一站完成沿 : Bool;
      扫码器接收数据 : String[16];
      扫码器扫码数值 : Int;
      扫码器扫码成功 : Bool;
   END_VAR
BEGIN
END_DATA_BLOCK

// folder: 通讯数据

DATA_BLOCK "虚拟联动信号"   // DB109
{ S7_Optimized_Access := 'FALSE' }
VERSION : 0.1
   VAR
      二站8mm挡停 : Bool;
      二站10mm挡停 : Bool;
      二站8mm推料 : Bool;
      二站10mm推料 : Bool;
      二站传送带 : Bool;
   END_VAR
BEGIN
END_DATA_BLOCK

DATA_BLOCK "一站数据"   // DB111
{ S7_Optimized_Access := 'FALSE' }
VERSION : 0.1
   VAR
      一站完成 : Bool;
      复位完成 : Bool;
      一站就绪 : Bool;
      一站忙碌 : Bool;
      一站请求二站接收 : Bool;
      一站可接单 : Bool;
      数据7 : Bool;
      数据8 : Bool;
      数据9 : Bool;
      数据10 : Bool;
      数据11 : Bool;
      数据12 : Bool;
      数据13 : Bool;
      数据14 : Bool;
   END_VAR
BEGIN
END_DATA_BLOCK

DATA_BLOCK "二站数据"   // DB112
{ S7_Optimized_Access := 'FALSE' }
VERSION : 0.1
   VAR
      二站完成 : Bool;
      二站已接收 : Bool;
      复位完成 : Bool;
      空闲状态 : Bool;
      电机正转 : Bool;
      二站忙碌 : Bool;
      二站请求三站接收 : Bool;
      二站可接收 : Bool;
      数据17 : Bool;
      数据18 : Bool;
      数据19 : Bool;
      数据20 : Bool;
      数据21 : Bool;
   END_VAR
BEGIN
END_DATA_BLOCK

DATA_BLOCK "三站数据"   // DB113
{ S7_Optimized_Access := 'FALSE' }
VERSION : 0.1
   VAR
      三站完成 : Bool;
      三站已接收 : Bool;
      复位完成 : Bool;
      空闲状态 : Bool;
      出现废料 : Bool;
      安全光栅 : Bool;
      三站可接收 : Bool;
      三站忙碌 : Bool;
      数据23 : Bool;
      数据24 : Bool;
      数据25 : Bool;
      数据26 : Bool;
      数据27 : Bool;
      数据28 : Bool;
      数据29 : Bool;
   END_VAR
BEGIN
END_DATA_BLOCK

DATA_BLOCK "AI视觉信号映射数据"   // DB116
{ S7_Optimized_Access := 'FALSE' }
VERSION : 0.1
   VAR
      二站上料完成 : Bool;
      钢珠灌料完成 : Bool;
   END_VAR
BEGIN
END_DATA_BLOCK

// folder: (top level)

FUNCTION "0.初始化" : Void   // FC1, LAD
{ S7_Optimized_Access := 'TRUE' }
VERSION : 0.1
   VAR_TEMP   // added for the SCL form of the ladder/FBD networks
      _w1 : Bool;
      _w2 : Bool;
   END_VAR
BEGIN

REGION Network 1: 模式切换
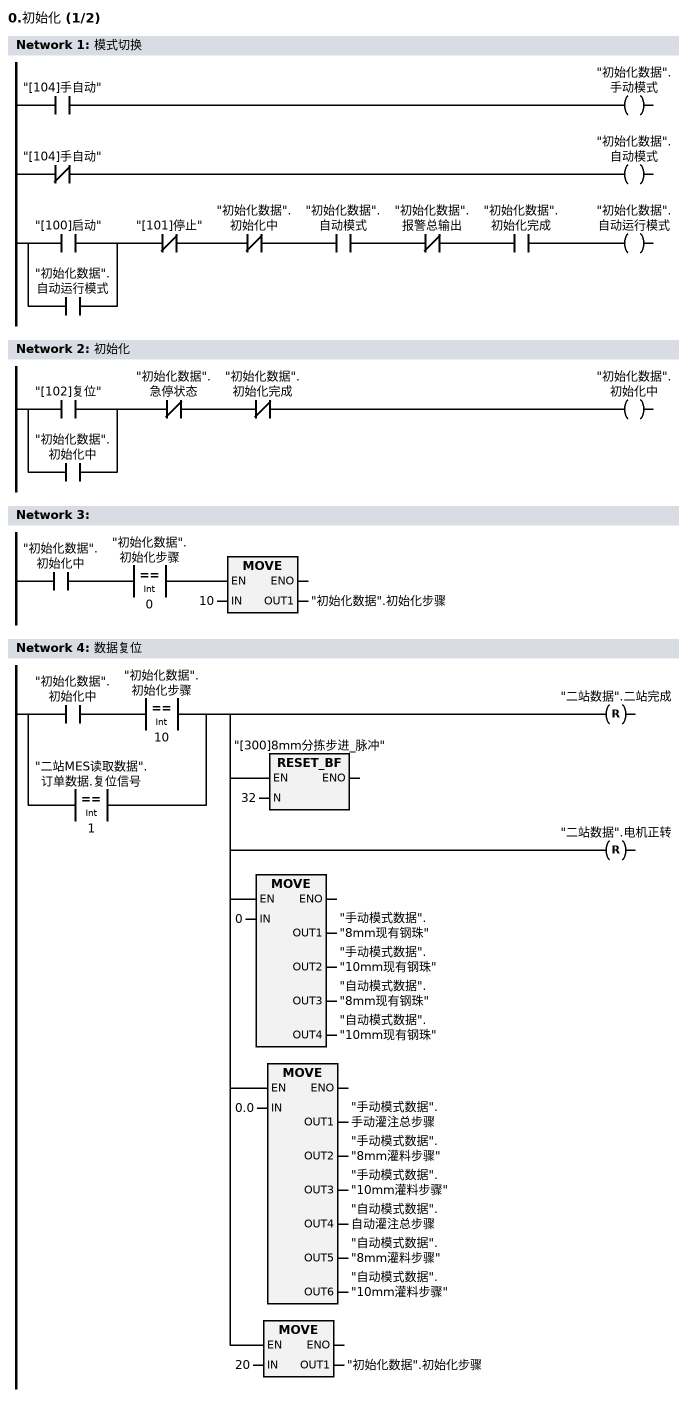
   RUNG wire#powerrail
      Contact( "[104]手自动" )
      Coil( "初始化数据".手动模式 )
   END_RUNG
   RUNG wire#powerrail
      I_Contact( "[104]手自动" )
      Coil( "初始化数据".自动模式 )
   END_RUNG
   RUNG wire#powerrail
      Contact( "[100]启动" )
      wire#w1
      I_Contact( "[101]停止" )
      I_Contact( "初始化数据".初始化中 )
      Contact( "初始化数据".自动模式 )
      I_Contact( "初始化数据".报警总输出 )
      Contact( "初始化数据".初始化完成 )
      Coil( "初始化数据".自动运行模式 )
   END_RUNG
   RUNG wire#powerrail
      Contact( "初始化数据".自动运行模式 )
   END_RUNG wire#w1
   // the same network as SCL:
   "初始化数据".手动模式 := "[104]手自动";
   "初始化数据".自动模式 := NOT "[104]手自动";
   "初始化数据".自动运行模式 := ("[100]启动" OR "初始化数据".自动运行模式) AND NOT "[101]停止" AND NOT "初始化数据".初始化中 AND "初始化数据".自动模式 AND NOT "初始化数据".报警总输出 AND "初始化数据".初始化完成;
END_REGION

REGION Network 2: 初始化
   RUNG wire#powerrail
      Contact( "[102]复位" )
      wire#w1
      I_Contact( "初始化数据".急停状态 )
      I_Contact( "初始化数据".初始化完成 )
      Coil( "初始化数据".初始化中 )
   END_RUNG
   RUNG wire#powerrail
      Contact( "初始化数据".初始化中 )
   END_RUNG wire#w1
   // the same network as SCL:
   "初始化数据".初始化中 := ("[102]复位" OR "初始化数据".初始化中) AND NOT "初始化数据".急停状态 AND NOT "初始化数据".初始化完成;
END_REGION

REGION Network 3
   RUNG wire#powerrail
      Contact( "初始化数据".初始化中 )
      { S7_Templates := "SrcType := Int" } EQ_Contact(in1 := "初始化数据".初始化步骤, in2 := 0)
      Move(in := 10, out1 => "初始化数据".初始化步骤)
   END_RUNG
   // the same network as SCL:
   IF "初始化数据".初始化中 AND ("初始化数据".初始化步骤 = 0) THEN "初始化数据".初始化步骤 := 10; END_IF;
END_REGION

REGION Network 4: 数据复位
   // no SCL statement known for RBitfield: written as a call
   IF ("初始化数据".初始化中 AND ("初始化数据".初始化步骤 = 10)) OR ("二站MES读取数据".订单数据.复位信号 = 1) THEN
       "二站数据".二站完成 := FALSE;
   END_IF;
   #_w1 := ("初始化数据".初始化中 AND ("初始化数据".初始化步骤 = 10)) OR ("二站MES读取数据".订单数据.复位信号 = 1);
   IF #_w1 THEN
       RESET_BF(operand := "[300]8mm分拣步进_脉冲", n := 32);
       "二站数据".电机正转 := FALSE;
       "手动模式数据"."8mm现有钢珠" := 0;
       "手动模式数据"."10mm现有钢珠" := 0;
       "自动模式数据"."8mm现有钢珠" := 0;
       "自动模式数据"."10mm现有钢珠" := 0;
       "手动模式数据".手动灌注总步骤 := 0.0;
       "手动模式数据"."8mm灌料步骤" := 0.0;
       "手动模式数据"."10mm灌料步骤" := 0.0;
       "自动模式数据".自动灌注总步骤 := 0.0;
       "自动模式数据"."8mm灌料步骤" := 0.0;
       "自动模式数据"."10mm灌料步骤" := 0.0;
       "初始化数据".初始化步骤 := 20;
   END_IF;
END_REGION

REGION Network 5: 初始化完成
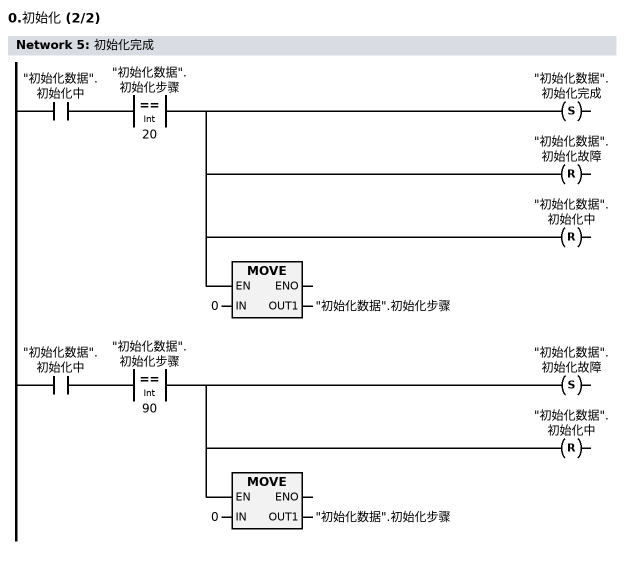
   RUNG wire#powerrail
      Contact( "初始化数据".初始化中 )
      { S7_Templates := "SrcType := Int" } EQ_Contact(in1 := "初始化数据".初始化步骤, in2 := 20)
      wire#w1
      S_Coil( "初始化数据".初始化完成 )
   END_RUNG
   RUNG wire#w1
      R_Coil( "初始化数据".初始化故障 )
   END_RUNG
   RUNG wire#w1
      R_Coil( "初始化数据".初始化中 )
   END_RUNG
   RUNG wire#w1
      Move(in := 0, out1 => "初始化数据".初始化步骤)
   END_RUNG
   RUNG wire#powerrail
      Contact( "初始化数据".初始化中 )
      { S7_Templates := "SrcType := Int" } EQ_Contact(in1 := "初始化数据".初始化步骤, in2 := 90)
      wire#w2
      S_Coil( "初始化数据".初始化故障 )
   END_RUNG
   RUNG wire#w2
      R_Coil( "初始化数据".初始化中 )
   END_RUNG
   RUNG wire#w2
      Move(in := 0, out1 => "初始化数据".初始化步骤)
   END_RUNG
   // the same network as SCL:
   IF "初始化数据".初始化中 AND ("初始化数据".初始化步骤 = 20) THEN
       "初始化数据".初始化完成 := TRUE;
       "初始化数据".初始化故障 := FALSE;
   END_IF;
   #_w1 := "初始化数据".初始化中 AND ("初始化数据".初始化步骤 = 20);
   IF #_w1 THEN
       "初始化数据".初始化中 := FALSE;
       "初始化数据".初始化步骤 := 0;
   END_IF;
   IF "初始化数据".初始化中 AND ("初始化数据".初始化步骤 = 90) THEN "初始化数据".初始化故障 := TRUE; END_IF;
   #_w2 := "初始化数据".初始化中 AND ("初始化数据".初始化步骤 = 90);
   IF #_w2 THEN
       "初始化数据".初始化中 := FALSE;
       "初始化数据".初始化步骤 := 0;
   END_IF;
END_REGION
END_FUNCTION

FUNCTION "2.状态控制" : Void   // FC9, LAD
{ S7_Optimized_Access := 'TRUE' }
VERSION : 0.1
BEGIN

REGION Network 1: 二站四种状态判断
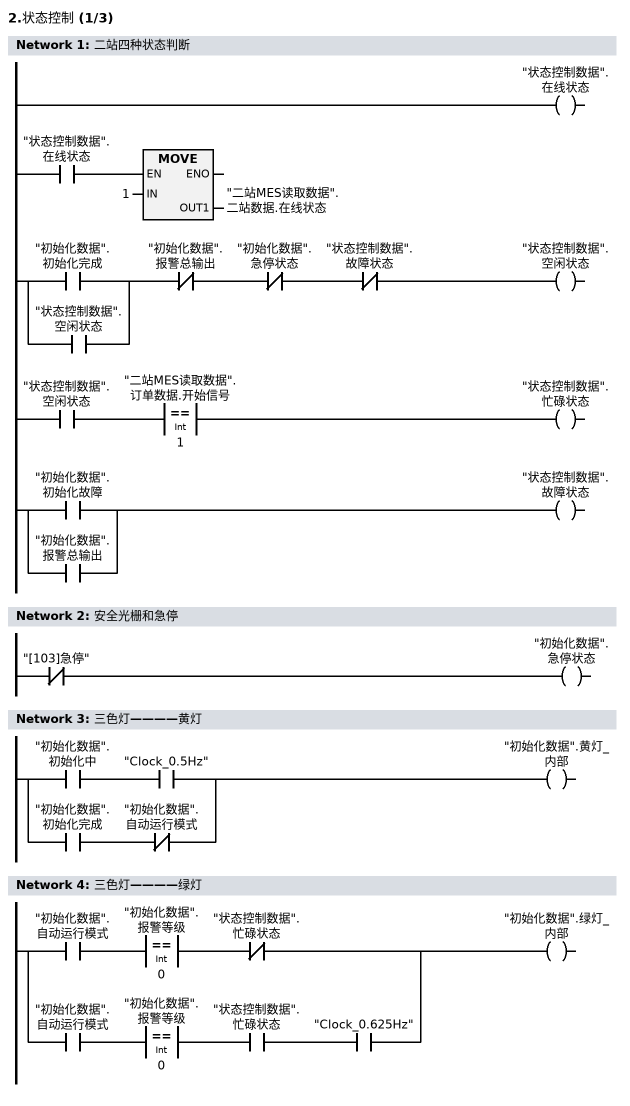
   RUNG wire#powerrail
      Coil( "状态控制数据".在线状态 )
   END_RUNG
   RUNG wire#powerrail
      Contact( "状态控制数据".在线状态 )
      Move(in := 1, out1 => "二站MES读取数据".二站数据.在线状态)
   END_RUNG
   RUNG wire#powerrail
      Contact( "初始化数据".初始化完成 )
      wire#w1
      I_Contact( "初始化数据".报警总输出 )
      I_Contact( "初始化数据".急停状态 )
      I_Contact( "状态控制数据".故障状态 )
      Coil( "状态控制数据".空闲状态 )
   END_RUNG
   RUNG wire#powerrail
      Contact( "状态控制数据".空闲状态 )
   END_RUNG wire#w1
   RUNG wire#powerrail
      Contact( "状态控制数据".空闲状态 )
      { S7_Templates := "SrcType := Int" } EQ_Contact(in1 := "二站MES读取数据".订单数据.开始信号, in2 := 1)
      Coil( "状态控制数据".忙碌状态 )
   END_RUNG
   RUNG wire#powerrail
      Contact( "初始化数据".初始化故障 )
      wire#w2
      Coil( "状态控制数据".故障状态 )
   END_RUNG
   RUNG wire#powerrail
      Contact( "初始化数据".报警总输出 )
   END_RUNG wire#w2
   // the same network as SCL:
   "状态控制数据".在线状态 := TRUE;
   IF "状态控制数据".在线状态 THEN "二站MES读取数据".二站数据.在线状态 := 1; END_IF;
   "状态控制数据".空闲状态 := ("初始化数据".初始化完成 OR "状态控制数据".空闲状态) AND NOT "初始化数据".报警总输出 AND NOT "初始化数据".急停状态 AND NOT "状态控制数据".故障状态;
   "状态控制数据".忙碌状态 := "状态控制数据".空闲状态 AND ("二站MES读取数据".订单数据.开始信号 = 1);
   "状态控制数据".故障状态 := "初始化数据".初始化故障 OR "初始化数据".报警总输出;
END_REGION

REGION Network 2: 安全光栅和急停
   RUNG wire#powerrail
      I_Contact( "[103]急停" )
      Coil( "初始化数据".急停状态 )
   END_RUNG
   // the same network as SCL:
   "初始化数据".急停状态 := NOT "[103]急停";
END_REGION

REGION Network 3: 三色灯————黄灯
   RUNG wire#powerrail
      Contact( "初始化数据".初始化中 )
      Contact( "Clock_0.5Hz" )
      wire#w1
      Coil( "初始化数据".黄灯_内部 )
   END_RUNG
   RUNG wire#powerrail
      Contact( "初始化数据".初始化完成 )
      I_Contact( "初始化数据".自动运行模式 )
   END_RUNG wire#w1
   // the same network as SCL:
   "初始化数据".黄灯_内部 := ("初始化数据".初始化中 AND "Clock_0.5Hz") OR ("初始化数据".初始化完成 AND NOT "初始化数据".自动运行模式);
END_REGION

REGION Network 4: 三色灯————绿灯
   RUNG wire#powerrail
      Contact( "初始化数据".自动运行模式 )
      { S7_Templates := "SrcType := Int" } EQ_Contact(in1 := "初始化数据".报警等级, in2 := 0)
      I_Contact( "状态控制数据".忙碌状态 )
      wire#w1
      Coil( "初始化数据".绿灯_内部 )
   END_RUNG
   RUNG wire#powerrail
      Contact( "初始化数据".自动运行模式 )
      { S7_Templates := "SrcType := Int" } EQ_Contact(in1 := "初始化数据".报警等级, in2 := 0)
      Contact( "状态控制数据".忙碌状态 )
      Contact( "Clock_0.625Hz" )
   END_RUNG wire#w1
   // the same network as SCL:
   "初始化数据".绿灯_内部 := ("初始化数据".自动运行模式 AND ("初始化数据".报警等级 = 0) AND NOT "状态控制数据".忙碌状态) OR ("初始化数据".自动运行模式 AND ("初始化数据".报警等级 = 0) AND "状态控制数据".忙碌状态 AND "Clock_0.625Hz");
END_REGION

REGION Network 5: 三色灯————红灯
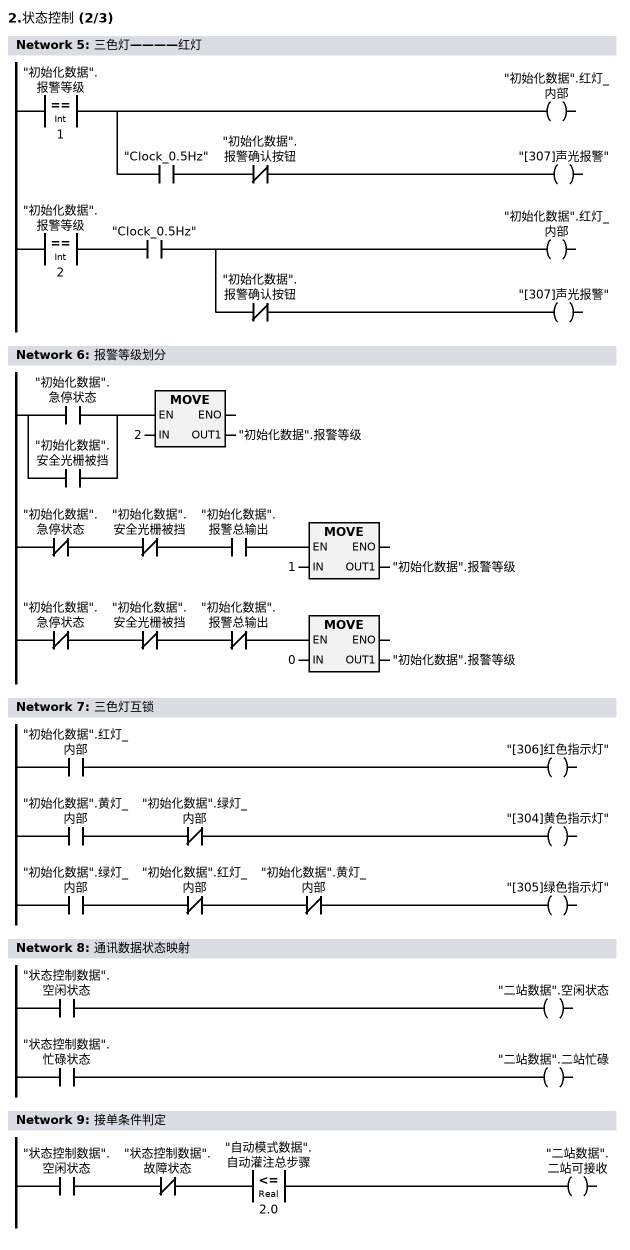
   RUNG wire#powerrail
      { S7_Templates := "SrcType := Int" } EQ_Contact(in1 := "初始化数据".报警等级, in2 := 1)
      wire#w1
      Coil( "初始化数据".红灯_内部 )
   END_RUNG
   RUNG wire#w1
      Contact( "Clock_0.5Hz" )
      I_Contact( "初始化数据".报警确认按钮 )
      Coil( "[307]声光报警" )
   END_RUNG
   RUNG wire#powerrail
      { S7_Templates := "SrcType := Int" } EQ_Contact(in1 := "初始化数据".报警等级, in2 := 2)
      Contact( "Clock_0.5Hz" )
      wire#w2
      Coil( "初始化数据".红灯_内部 )
   END_RUNG
   RUNG wire#w2
      I_Contact( "初始化数据".报警确认按钮 )
      Coil( "[307]声光报警" )
   END_RUNG
   // the same network as SCL:
   "初始化数据".红灯_内部 := "初始化数据".报警等级 = 1;
   "[307]声光报警" := "初始化数据".红灯_内部 AND "Clock_0.5Hz" AND NOT "初始化数据".报警确认按钮;
   "初始化数据".红灯_内部 := ("初始化数据".报警等级 = 2) AND "Clock_0.5Hz";
   "[307]声光报警" := "初始化数据".红灯_内部 AND NOT "初始化数据".报警确认按钮;
END_REGION

REGION Network 6: 报警等级划分
   RUNG wire#powerrail
      Contact( "初始化数据".急停状态 )
      wire#w1
      Move(in := 2, out1 => "初始化数据".报警等级)
   END_RUNG
   RUNG wire#powerrail
      Contact( "初始化数据".安全光栅被挡 )
   END_RUNG wire#w1
   RUNG wire#powerrail
      I_Contact( "初始化数据".急停状态 )
      I_Contact( "初始化数据".安全光栅被挡 )
      Contact( "初始化数据".报警总输出 )
      Move(in := 1, out1 => "初始化数据".报警等级)
   END_RUNG
   RUNG wire#powerrail
      I_Contact( "初始化数据".急停状态 )
      I_Contact( "初始化数据".安全光栅被挡 )
      I_Contact( "初始化数据".报警总输出 )
      Move(in := 0, out1 => "初始化数据".报警等级)
   END_RUNG
   // the same network as SCL:
   IF "初始化数据".急停状态 OR "初始化数据".安全光栅被挡 THEN "初始化数据".报警等级 := 2; END_IF;
   IF NOT "初始化数据".急停状态 AND NOT "初始化数据".安全光栅被挡 AND "初始化数据".报警总输出 THEN "初始化数据".报警等级 := 1; END_IF;
   IF NOT "初始化数据".急停状态 AND NOT "初始化数据".安全光栅被挡 AND NOT "初始化数据".报警总输出 THEN "初始化数据".报警等级 := 0; END_IF;
END_REGION

REGION Network 7: 三色灯互锁
   RUNG wire#powerrail
      Contact( "初始化数据".红灯_内部 )
      Coil( "[306]红色指示灯" )
   END_RUNG
   RUNG wire#powerrail
      Contact( "初始化数据".黄灯_内部 )
      I_Contact( "初始化数据".绿灯_内部 )
      Coil( "[304]黄色指示灯" )
   END_RUNG
   RUNG wire#powerrail
      Contact( "初始化数据".绿灯_内部 )
      I_Contact( "初始化数据".红灯_内部 )
      I_Contact( "初始化数据".黄灯_内部 )
      Coil( "[305]绿色指示灯" )
   END_RUNG
   // the same network as SCL:
   "[306]红色指示灯" := "初始化数据".红灯_内部;
   "[304]黄色指示灯" := "初始化数据".黄灯_内部 AND NOT "初始化数据".绿灯_内部;
   "[305]绿色指示灯" := "初始化数据".绿灯_内部 AND NOT "初始化数据".红灯_内部 AND NOT "初始化数据".黄灯_内部;
END_REGION

REGION Network 8: 通讯数据状态映射
   RUNG wire#powerrail
      Contact( "状态控制数据".空闲状态 )
      Coil( "二站数据".空闲状态 )
   END_RUNG
   RUNG wire#powerrail
      Contact( "状态控制数据".忙碌状态 )
      Coil( "二站数据".二站忙碌 )
   END_RUNG
   // the same network as SCL:
   "二站数据".空闲状态 := "状态控制数据".空闲状态;
   "二站数据".二站忙碌 := "状态控制数据".忙碌状态;
END_REGION

REGION Network 9: 接单条件判定
   RUNG wire#powerrail
      Contact( "状态控制数据".空闲状态 )
      I_Contact( "状态控制数据".故障状态 )
      { S7_Templates := "SrcType := Real" } LE_Contact(in1 := "自动模式数据".自动灌注总步骤, in2 := 2.0)
      Coil( "二站数据".二站可接收 )
   END_RUNG
   // the same network as SCL:
   "二站数据".二站可接收 := "状态控制数据".空闲状态 AND NOT "状态控制数据".故障状态 AND ("自动模式数据".自动灌注总步骤 <= 2.0);
END_REGION

REGION Network 10: MES通讯映射
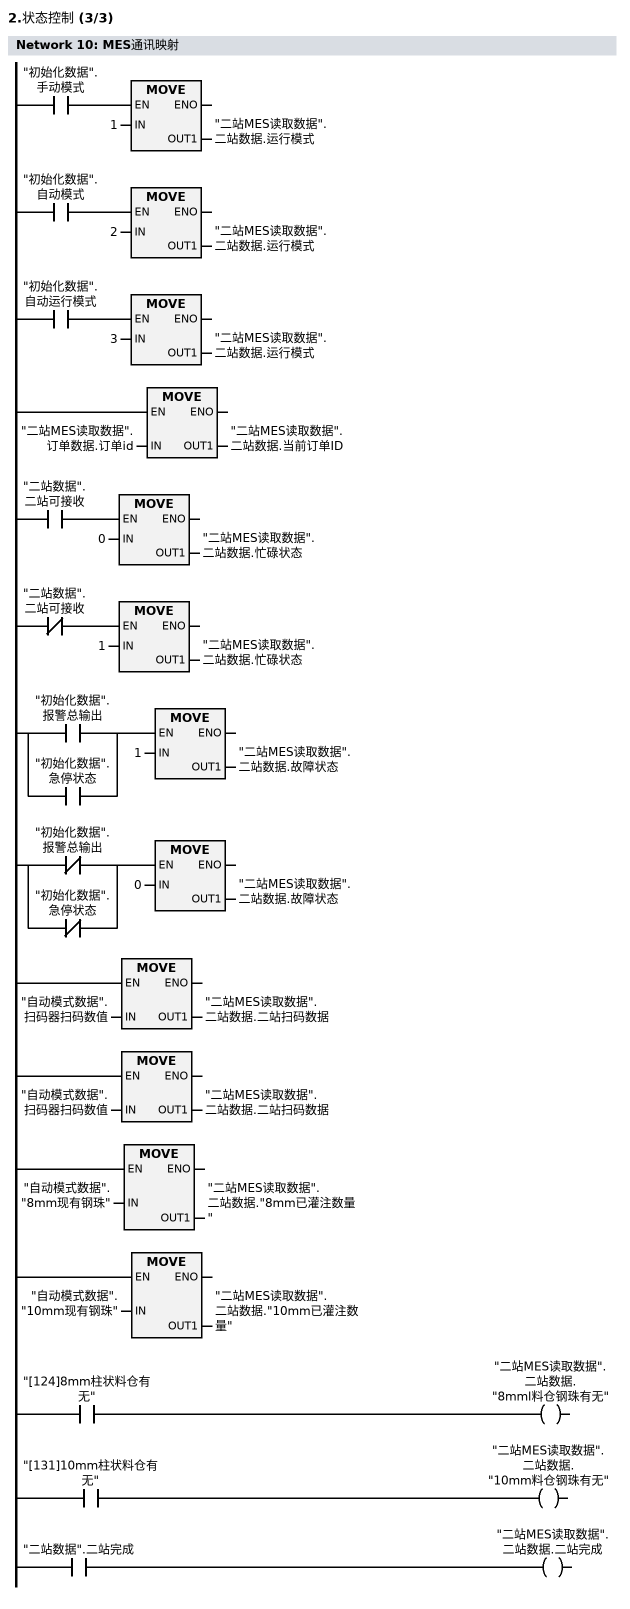
   RUNG wire#powerrail
      Contact( "初始化数据".手动模式 )
      Move(in := 1, out1 => "二站MES读取数据".二站数据.运行模式)
   END_RUNG
   RUNG wire#powerrail
      Contact( "初始化数据".自动模式 )
      Move(in := 2, out1 => "二站MES读取数据".二站数据.运行模式)
   END_RUNG
   RUNG wire#powerrail
      Contact( "初始化数据".自动运行模式 )
      Move(in := 3, out1 => "二站MES读取数据".二站数据.运行模式)
   END_RUNG
   RUNG wire#powerrail
      Move(in := "二站MES读取数据".订单数据.订单id, out1 => "二站MES读取数据".二站数据.当前订单ID)
   END_RUNG
   RUNG wire#powerrail
      Contact( "二站数据".二站可接收 )
      Move(in := 0, out1 => "二站MES读取数据".二站数据.忙碌状态)
   END_RUNG
   RUNG wire#powerrail
      I_Contact( "二站数据".二站可接收 )
      Move(in := 1, out1 => "二站MES读取数据".二站数据.忙碌状态)
   END_RUNG
   RUNG wire#powerrail
      Contact( "初始化数据".报警总输出 )
      wire#w1
      Move(in := 1, out1 => "二站MES读取数据".二站数据.故障状态)
   END_RUNG
   RUNG wire#powerrail
      Contact( "初始化数据".急停状态 )
   END_RUNG wire#w1
   RUNG wire#powerrail
      I_Contact( "初始化数据".报警总输出 )
      wire#w2
      Move(in := 0, out1 => "二站MES读取数据".二站数据.故障状态)
   END_RUNG
   RUNG wire#powerrail
      I_Contact( "初始化数据".急停状态 )
   END_RUNG wire#w2
   RUNG wire#powerrail
      Move(in := "自动模式数据".扫码器扫码数值, out1 => "二站MES读取数据".二站数据.二站扫码数据)
   END_RUNG
   RUNG wire#powerrail
      Move(in := "自动模式数据".扫码器扫码数值, out1 => "二站MES读取数据".二站数据.二站扫码数据)
   END_RUNG
   RUNG wire#powerrail
      Move(in := "自动模式数据"."8mm现有钢珠", out1 => "二站MES读取数据".二站数据."8mm已灌注数量")
   END_RUNG
   RUNG wire#powerrail
      Move(in := "自动模式数据"."10mm现有钢珠", out1 => "二站MES读取数据".二站数据."10mm已灌注数量")
   END_RUNG
   RUNG wire#powerrail
      Contact( "[124]8mm柱状料仓有无" )
      Coil( "二站MES读取数据".二站数据."8mml料仓钢珠有无" )
   END_RUNG
   RUNG wire#powerrail
      Contact( "[131]10mm柱状料仓有无" )
      Coil( "二站MES读取数据".二站数据."10mm料仓钢珠有无" )
   END_RUNG
   RUNG wire#powerrail
      Contact( "二站数据".二站完成 )
      Coil( "二站MES读取数据".二站数据.二站完成 )
   END_RUNG
   // the same network as SCL:
   IF "初始化数据".手动模式 THEN "二站MES读取数据".二站数据.运行模式 := 1; END_IF;
   IF "初始化数据".自动模式 THEN "二站MES读取数据".二站数据.运行模式 := 2; END_IF;
   IF "初始化数据".自动运行模式 THEN "二站MES读取数据".二站数据.运行模式 := 3; END_IF;
   "二站MES读取数据".二站数据.当前订单ID := "二站MES读取数据".订单数据.订单id;
   IF "二站数据".二站可接收 THEN "二站MES读取数据".二站数据.忙碌状态 := 0; END_IF;
   IF NOT "二站数据".二站可接收 THEN "二站MES读取数据".二站数据.忙碌状态 := 1; END_IF;
   IF "初始化数据".报警总输出 OR "初始化数据".急停状态 THEN "二站MES读取数据".二站数据.故障状态 := 1; END_IF;
   IF NOT "初始化数据".报警总输出 OR NOT "初始化数据".急停状态 THEN "二站MES读取数据".二站数据.故障状态 := 0; END_IF;
   "二站MES读取数据".二站数据.二站扫码数据 := "自动模式数据".扫码器扫码数值;
   "二站MES读取数据".二站数据.二站扫码数据 := "自动模式数据".扫码器扫码数值;
   "二站MES读取数据".二站数据."8mm已灌注数量" := "自动模式数据"."8mm现有钢珠";
   "二站MES读取数据".二站数据."10mm已灌注数量" := "自动模式数据"."10mm现有钢珠";
   "二站MES读取数据".二站数据."8mml料仓钢珠有无" := "[124]8mm柱状料仓有无";
   "二站MES读取数据".二站数据."10mm料仓钢珠有无" := "[131]10mm柱状料仓有无";
   "二站MES读取数据".二站数据.二站完成 := "二站数据".二站完成;
END_REGION
END_FUNCTION

FUNCTION "1.报警程序" : Void   // FC13, LAD
{ S7_Optimized_Access := 'TRUE' }
VERSION : 0.1
BEGIN

REGION Network 1: 气缸报警——————8mm挡停气缸
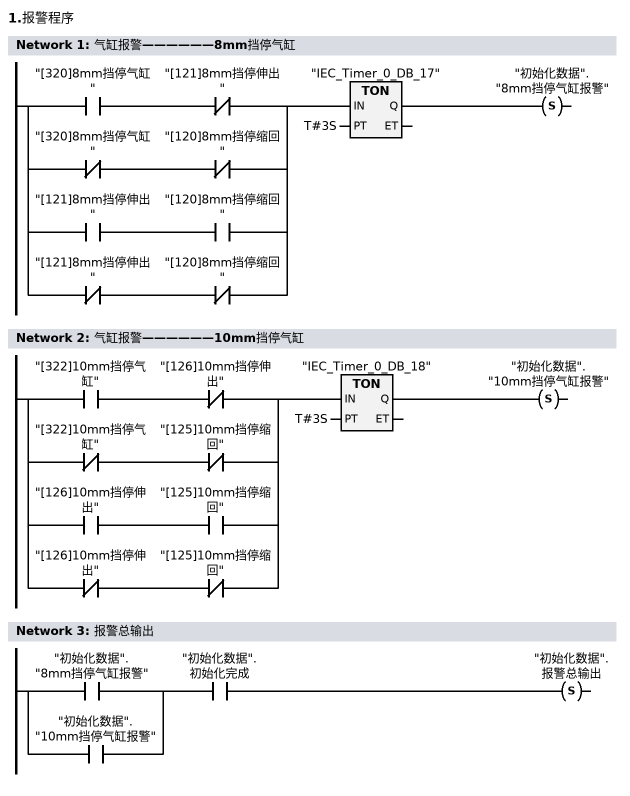
   "IEC_Timer_0_DB_17".TON(IN := ("[320]8mm挡停气缸" AND NOT "[121]8mm挡停伸出") OR (NOT "[320]8mm挡停气缸" AND NOT "[120]8mm挡停缩回") OR ("[121]8mm挡停伸出" AND "[120]8mm挡停缩回") OR (NOT "[121]8mm挡停伸出" AND NOT "[120]8mm挡停缩回"),
                           PT := T#3S);
   IF "IEC_Timer_0_DB_17".Q THEN "初始化数据"."8mm挡停气缸报警" := TRUE; END_IF;
END_REGION

REGION Network 2: 气缸报警——————10mm挡停气缸
   "IEC_Timer_0_DB_18".TON(IN := ("[322]10mm挡停气缸" AND NOT "[126]10mm挡停伸出") OR (NOT "[322]10mm挡停气缸" AND NOT "[125]10mm挡停缩回") OR ("[126]10mm挡停伸出" AND "[125]10mm挡停缩回") OR (NOT "[126]10mm挡停伸出" AND NOT "[125]10mm挡停缩回"),
                           PT := T#3S);
   IF "IEC_Timer_0_DB_18".Q THEN "初始化数据"."10mm挡停气缸报警" := TRUE; END_IF;
END_REGION

REGION Network 3: 报警总输出
   RUNG wire#powerrail
      Contact( "初始化数据"."8mm挡停气缸报警" )
      wire#w1
      Contact( "初始化数据".初始化完成 )
      S_Coil( "初始化数据".报警总输出 )
   END_RUNG
   RUNG wire#powerrail
      Contact( "初始化数据"."10mm挡停气缸报警" )
   END_RUNG wire#w1
   // the same network as SCL:
   IF ("初始化数据"."8mm挡停气缸报警" OR "初始化数据"."10mm挡停气缸报警") AND "初始化数据".初始化完成 THEN "初始化数据".报警总输出 := TRUE; END_IF;
END_REGION

REGION Network 4: 触发声光报警
END_REGION
END_FUNCTION

ORGANIZATION_BLOCK "Main"   // OB1, LAD, ProgramCycle
TITLE = "Main Program Sweep (Cycle)"
{ S7_Optimized_Access := 'TRUE' }
VERSION : 0.1
   VAR_INPUT
      Initial_Call : Bool;   // Initial call of this OB
      Remanence : Bool;   // =True, if remanent data are available
   END_VAR
   VAR_TEMP   // added for the SCL form of the ladder/FBD networks
      _w1 : Bool;
      _w2 : Bool;
      _w3 : Bool;
      _w4 : Bool;
   END_VAR
BEGIN

REGION Network 1: 自动模式
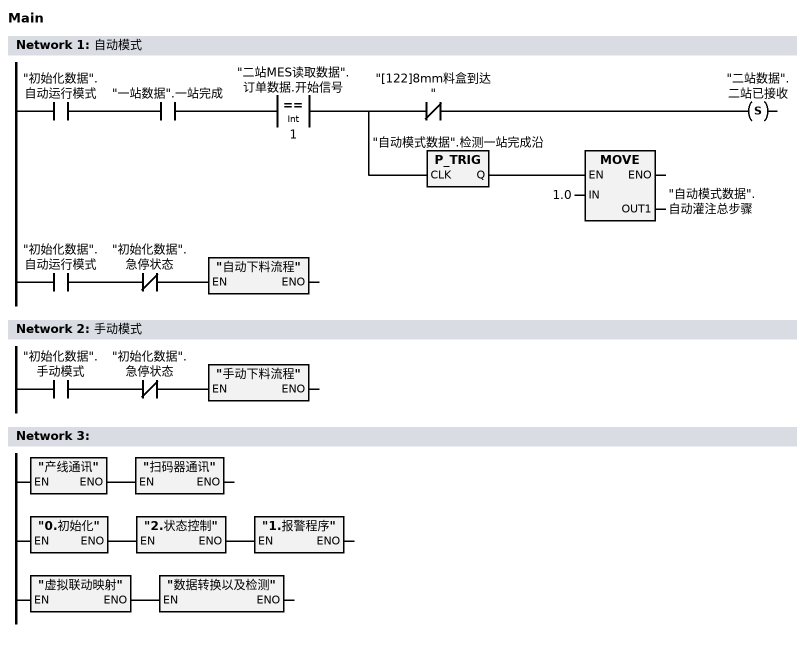
   RUNG wire#powerrail
      Contact( "初始化数据".自动运行模式 )
      Contact( "一站数据".一站完成 )
      { S7_Templates := "SrcType := Int" } EQ_Contact(in1 := "二站MES读取数据".订单数据.开始信号, in2 := 1)
      wire#w1
      I_Contact( "[122]8mm料盒到达" )
      S_Coil( "二站数据".二站已接收 )
   END_RUNG
   RUNG wire#w1
      P_Trig( "自动模式数据".检测一站完成沿 )
      Move(in := 1.0, out1 => "自动模式数据".自动灌注总步骤)
   END_RUNG
   RUNG wire#powerrail
      Contact( "初始化数据".自动运行模式 )
      I_Contact( "初始化数据".急停状态 )
      "自动下料流程"()
   END_RUNG
   // the same network as SCL:
   #_w1 := "初始化数据".自动运行模式 AND "一站数据".一站完成 AND ("二站MES读取数据".订单数据.开始信号 = 1);
   IF #_w1 AND NOT "[122]8mm料盒到达" THEN "二站数据".二站已接收 := TRUE; END_IF;
   #_w2 := #_w1 AND NOT "自动模式数据".检测一站完成沿;   // rising edge
   "自动模式数据".检测一站完成沿 := #_w1;
   IF #_w2 THEN "自动模式数据".自动灌注总步骤 := 1.0; END_IF;
   IF "初始化数据".自动运行模式 AND NOT "初始化数据".急停状态 THEN "自动下料流程"(); END_IF;
END_REGION

REGION Network 2: 手动模式
   RUNG wire#powerrail
      Contact( "初始化数据".手动模式 )
      I_Contact( "初始化数据".急停状态 )
      "手动下料流程"()
   END_RUNG
   // the same network as SCL:
   IF "初始化数据".手动模式 AND NOT "初始化数据".急停状态 THEN "手动下料流程"(); END_IF;
END_REGION

REGION Network 3
   RUNG wire#powerrail
      "产线通讯"()
      "扫码器通讯"()
   END_RUNG
   RUNG wire#powerrail
      "0.初始化"()
      "2.状态控制"()
      "1.报警程序"()
   END_RUNG
   RUNG wire#powerrail
      "虚拟联动映射"()
      "数据转换以及检测"()
   END_RUNG
   // the same network as SCL:
   "产线通讯"(ENO => #_w1);
   IF #_w1 THEN "扫码器通讯"(); END_IF;
   "0.初始化"(ENO => #_w2);
   "2.状态控制"(EN := #_w2, ENO => #_w3);
   IF #_w3 THEN "1.报警程序"(); END_IF;
   "虚拟联动映射"(ENO => #_w4);
   IF #_w4 THEN "数据转换以及检测"(); END_IF;
END_REGION
END_ORGANIZATION_BLOCK

// folder: 手动模式

FUNCTION "手动下料流程" : Void   // FC3, LAD
{ S7_Optimized_Access := 'TRUE' }
VERSION : 0.1
   VAR_TEMP   // added for the SCL form of the ladder/FBD networks
      _w1 : Bool;
   END_VAR
BEGIN

REGION Network 1: 复位
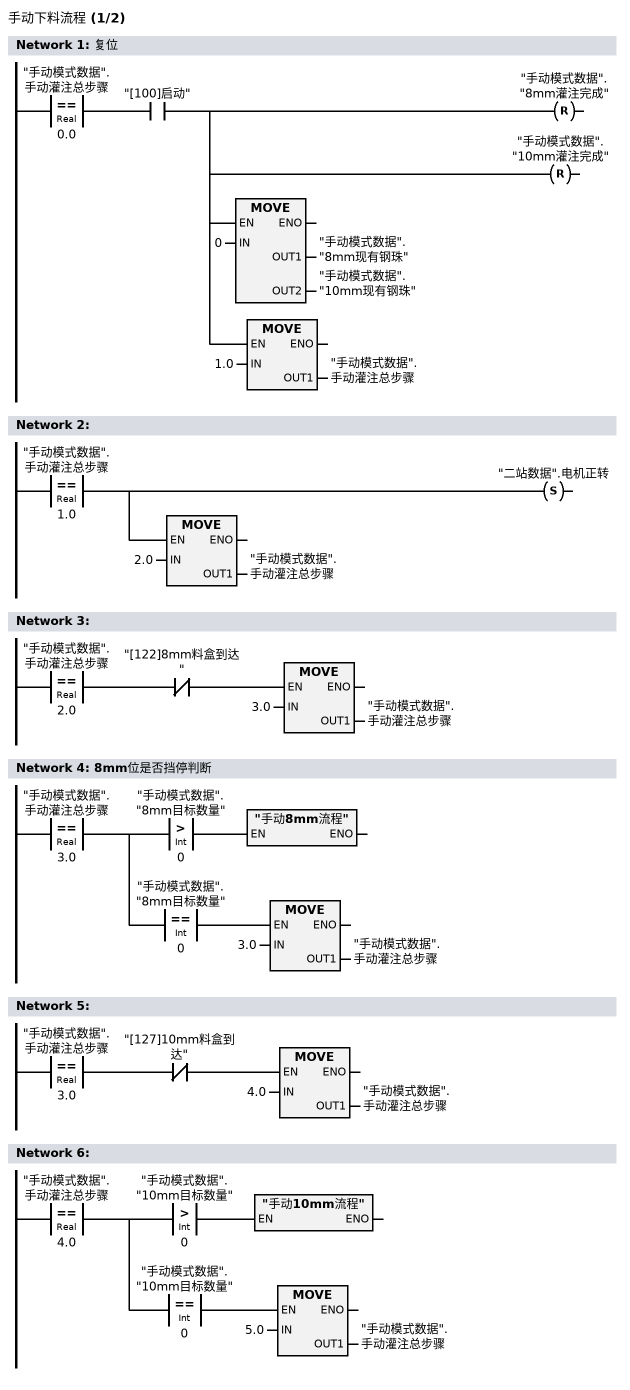
   RUNG wire#powerrail
      { S7_Templates := "SrcType := Real" } EQ_Contact(in1 := "手动模式数据".手动灌注总步骤, in2 := 0.0)
      Contact( "[100]启动" )
      wire#w1
      R_Coil( "手动模式数据"."8mm灌注完成" )
   END_RUNG
   RUNG wire#w1
      R_Coil( "手动模式数据"."10mm灌注完成" )
   END_RUNG
   RUNG wire#w1
      Move(in := 0, out1 => "手动模式数据"."8mm现有钢珠", out2 => "手动模式数据"."10mm现有钢珠")
   END_RUNG
   RUNG wire#w1
      Move(in := 1.0, out1 => "手动模式数据".手动灌注总步骤)
   END_RUNG
   // the same network as SCL:
   IF ("手动模式数据".手动灌注总步骤 = 0.0) AND "[100]启动" THEN
       "手动模式数据"."8mm灌注完成" := FALSE;
       "手动模式数据"."10mm灌注完成" := FALSE;
       "手动模式数据"."8mm现有钢珠" := 0;
       "手动模式数据"."10mm现有钢珠" := 0;
       "手动模式数据".手动灌注总步骤 := 1.0;
   END_IF;
END_REGION

REGION Network 2
   RUNG wire#powerrail
      { S7_Templates := "SrcType := Real" } EQ_Contact(in1 := "手动模式数据".手动灌注总步骤, in2 := 1.0)
      wire#w1
      S_Coil( "二站数据".电机正转 )
   END_RUNG
   RUNG wire#w1
      Move(in := 2.0, out1 => "手动模式数据".手动灌注总步骤)
   END_RUNG
   // the same network as SCL:
   IF "手动模式数据".手动灌注总步骤 = 1.0 THEN
       "二站数据".电机正转 := TRUE;
       "手动模式数据".手动灌注总步骤 := 2.0;
   END_IF;
END_REGION

REGION Network 3
   RUNG wire#powerrail
      { S7_Templates := "SrcType := Real" } EQ_Contact(in1 := "手动模式数据".手动灌注总步骤, in2 := 2.0)
      I_Contact( "[122]8mm料盒到达" )
      Move(in := 3.0, out1 => "手动模式数据".手动灌注总步骤)
   END_RUNG
   // the same network as SCL:
   IF ("手动模式数据".手动灌注总步骤 = 2.0) AND NOT "[122]8mm料盒到达" THEN "手动模式数据".手动灌注总步骤 := 3.0; END_IF;
END_REGION

REGION Network 4: 8mm位是否挡停判断
   RUNG wire#powerrail
      { S7_Templates := "SrcType := Real" } EQ_Contact(in1 := "手动模式数据".手动灌注总步骤, in2 := 3.0)
      wire#w1
      { S7_Templates := "SrcType := Int" } GT_Contact(in1 := "手动模式数据"."8mm目标数量", in2 := 0)
      "手动8mm流程"()
   END_RUNG
   RUNG wire#w1
      { S7_Templates := "SrcType := Int" } EQ_Contact(in1 := "手动模式数据"."8mm目标数量", in2 := 0)
      Move(in := 3.0, out1 => "手动模式数据".手动灌注总步骤)
   END_RUNG
   // the same network as SCL:
   #_w1 := "手动模式数据".手动灌注总步骤 = 3.0;
   IF #_w1 AND ("手动模式数据"."8mm目标数量" > 0) THEN "手动8mm流程"(); END_IF;
   IF #_w1 AND ("手动模式数据"."8mm目标数量" = 0) THEN "手动模式数据".手动灌注总步骤 := 3.0; END_IF;
END_REGION

REGION Network 5
   RUNG wire#powerrail
      { S7_Templates := "SrcType := Real" } EQ_Contact(in1 := "手动模式数据".手动灌注总步骤, in2 := 3.0)
      I_Contact( "[127]10mm料盒到达" )
      Move(in := 4.0, out1 => "手动模式数据".手动灌注总步骤)
   END_RUNG
   // the same network as SCL:
   IF ("手动模式数据".手动灌注总步骤 = 3.0) AND NOT "[127]10mm料盒到达" THEN "手动模式数据".手动灌注总步骤 := 4.0; END_IF;
END_REGION

REGION Network 6
   RUNG wire#powerrail
      { S7_Templates := "SrcType := Real" } EQ_Contact(in1 := "手动模式数据".手动灌注总步骤, in2 := 4.0)
      wire#w1
      { S7_Templates := "SrcType := Int" } GT_Contact(in1 := "手动模式数据"."10mm目标数量", in2 := 0)
      "手动10mm流程"()
   END_RUNG
   RUNG wire#w1
      { S7_Templates := "SrcType := Int" } EQ_Contact(in1 := "手动模式数据"."10mm目标数量", in2 := 0)
      Move(in := 5.0, out1 => "手动模式数据".手动灌注总步骤)
   END_RUNG
   // the same network as SCL:
   #_w1 := "手动模式数据".手动灌注总步骤 = 4.0;
   IF #_w1 AND ("手动模式数据"."10mm目标数量" > 0) THEN "手动10mm流程"(); END_IF;
   IF #_w1 AND ("手动模式数据"."10mm目标数量" = 0) THEN "手动模式数据".手动灌注总步骤 := 5.0; END_IF;
END_REGION

REGION Network 7: 输出完成信号，运输至第三站
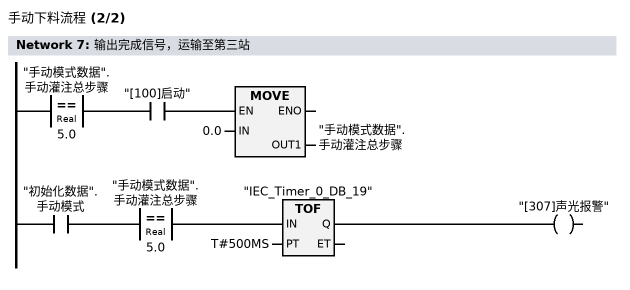
   IF ("手动模式数据".手动灌注总步骤 = 5.0) AND "[100]启动" THEN "手动模式数据".手动灌注总步骤 := 0.0; END_IF;
   "IEC_Timer_0_DB_19".TOF(IN := "初始化数据".手动模式 AND ("手动模式数据".手动灌注总步骤 = 5.0), PT := T#500MS);
   "[307]声光报警" := "IEC_Timer_0_DB_19".Q;
END_REGION
END_FUNCTION

FUNCTION "手动8mm流程" : Void   // FC4, LAD
{ S7_Optimized_Access := 'TRUE' }
VERSION : 0.1
   VAR_TEMP   // added for the SCL form of the ladder/FBD networks
      _w1 : Bool;
      _w2 : Bool;
   END_VAR
BEGIN

REGION Network 1
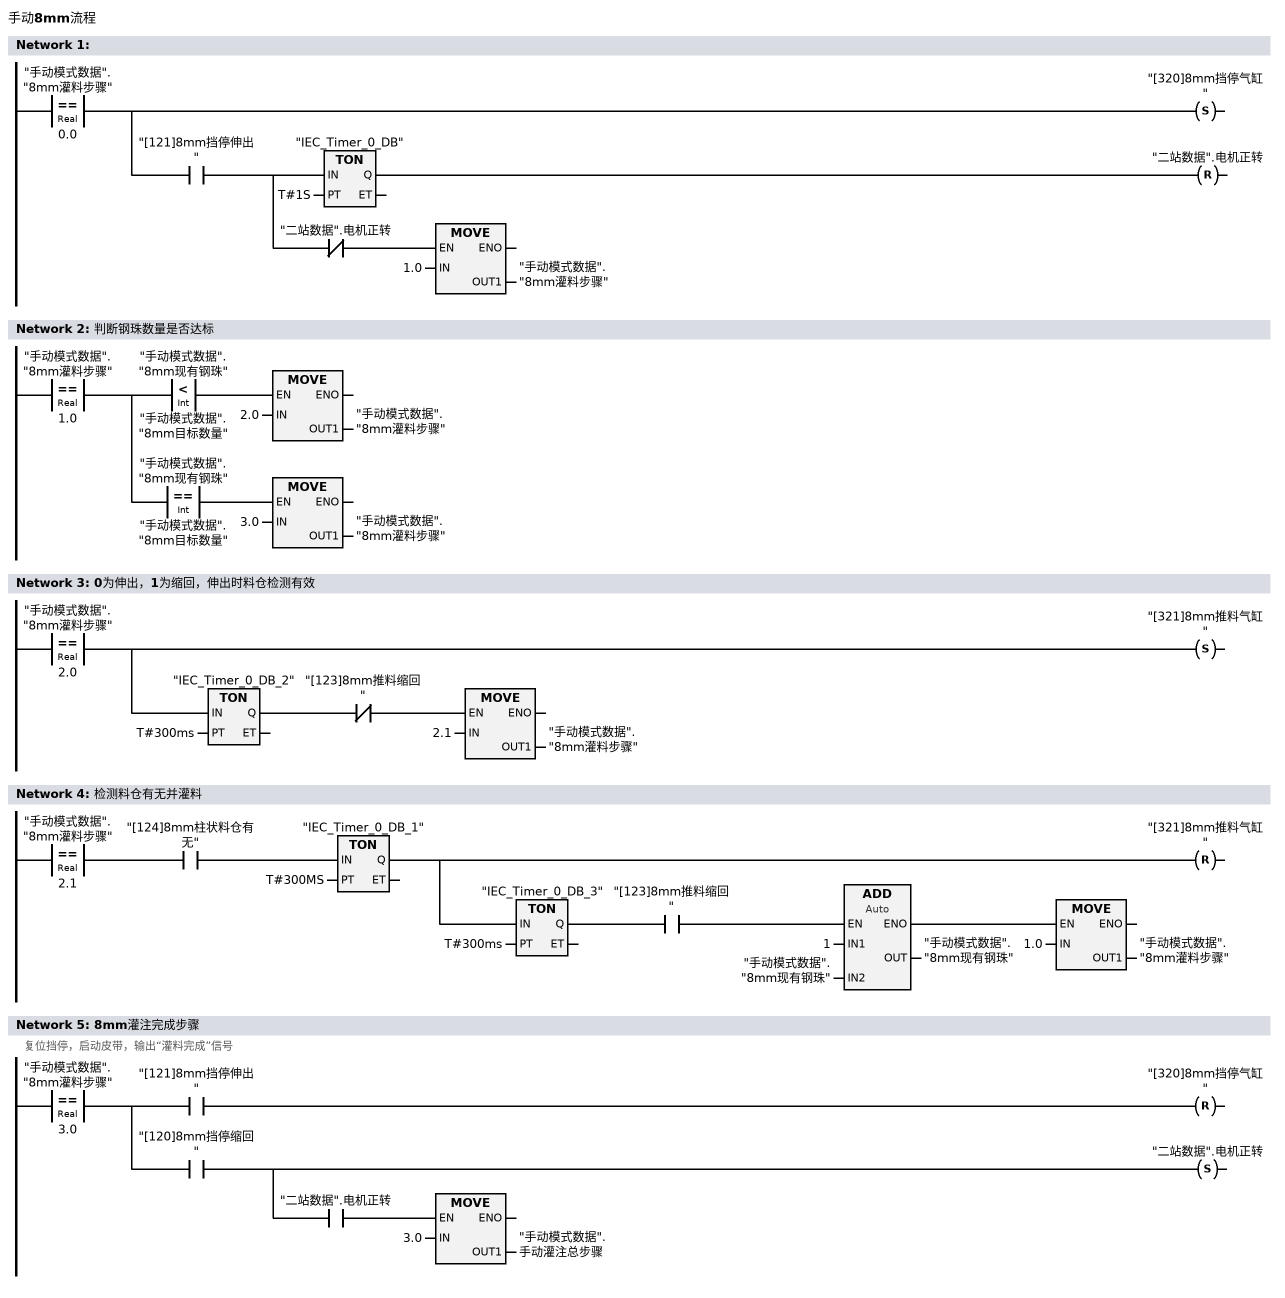
   #_w1 := "手动模式数据"."8mm灌料步骤" = 0.0;
   IF #_w1 THEN "[320]8mm挡停气缸" := TRUE; END_IF;
   #_w2 := #_w1 AND "[121]8mm挡停伸出";
   "IEC_Timer_0_DB".TON(IN := #_w2, PT := T#1S);
   IF "IEC_Timer_0_DB".Q THEN "二站数据".电机正转 := FALSE; END_IF;
   IF #_w2 AND NOT "二站数据".电机正转 THEN "手动模式数据"."8mm灌料步骤" := 1.0; END_IF;
END_REGION

REGION Network 2: 判断钢珠数量是否达标
   RUNG wire#powerrail
      { S7_Templates := "SrcType := Real" } EQ_Contact(in1 := "手动模式数据"."8mm灌料步骤", in2 := 1.0)
      wire#w1
      { S7_Templates := "SrcType := Int" } LT_Contact(in1 := "手动模式数据"."8mm现有钢珠", in2 := "手动模式数据"."8mm目标数量")
      Move(in := 2.0, out1 => "手动模式数据"."8mm灌料步骤")
   END_RUNG
   RUNG wire#w1
      { S7_Templates := "SrcType := Int" } EQ_Contact(in1 := "手动模式数据"."8mm现有钢珠", in2 := "手动模式数据"."8mm目标数量")
      Move(in := 3.0, out1 => "手动模式数据"."8mm灌料步骤")
   END_RUNG
   // the same network as SCL:
   #_w1 := "手动模式数据"."8mm灌料步骤" = 1.0;
   IF #_w1 AND ("手动模式数据"."8mm现有钢珠" < "手动模式数据"."8mm目标数量") THEN "手动模式数据"."8mm灌料步骤" := 2.0; END_IF;
   IF #_w1 AND ("手动模式数据"."8mm现有钢珠" = "手动模式数据"."8mm目标数量") THEN "手动模式数据"."8mm灌料步骤" := 3.0; END_IF;
END_REGION

REGION Network 3: 0为伸出，1为缩回，伸出时料仓检测有效
   #_w1 := "手动模式数据"."8mm灌料步骤" = 2.0;
   IF #_w1 THEN "[321]8mm推料气缸" := TRUE; END_IF;
   "IEC_Timer_0_DB_2".TON(IN := #_w1, PT := T#300ms);
   IF "IEC_Timer_0_DB_2".Q AND NOT "[123]8mm推料缩回" THEN "手动模式数据"."8mm灌料步骤" := 2.1; END_IF;
END_REGION

REGION Network 4: 检测料仓有无并灌料
   "IEC_Timer_0_DB_1".TON(IN := ("手动模式数据"."8mm灌料步骤" = 2.1) AND "[124]8mm柱状料仓有无", PT := T#300MS);
   IF "IEC_Timer_0_DB_1".Q THEN "[321]8mm推料气缸" := FALSE; END_IF;
   "IEC_Timer_0_DB_3".TON(IN := "IEC_Timer_0_DB_1".Q, PT := T#300ms);
   IF "IEC_Timer_0_DB_3".Q AND "[123]8mm推料缩回" THEN
       "手动模式数据"."8mm现有钢珠" := 1 + "手动模式数据"."8mm现有钢珠";
       "手动模式数据"."8mm灌料步骤" := 1.0;
   END_IF;
END_REGION

REGION Network 5: 8mm灌注完成步骤
   // 复位挡停，启动皮带，输出“灌料完成”信号
   RUNG wire#powerrail
      { S7_Templates := "SrcType := Real" } EQ_Contact(in1 := "手动模式数据"."8mm灌料步骤", in2 := 3.0)
      wire#w1
      Contact( "[121]8mm挡停伸出" )
      R_Coil( "[320]8mm挡停气缸" )
   END_RUNG
   RUNG wire#w1
      Contact( "[120]8mm挡停缩回" )
      wire#w2
      S_Coil( "二站数据".电机正转 )
   END_RUNG
   RUNG wire#w2
      Contact( "二站数据".电机正转 )
      Move(in := 3.0, out1 => "手动模式数据".手动灌注总步骤)
   END_RUNG
   // the same network as SCL:
   #_w1 := "手动模式数据"."8mm灌料步骤" = 3.0;
   IF #_w1 AND "[121]8mm挡停伸出" THEN "[320]8mm挡停气缸" := FALSE; END_IF;
   #_w2 := #_w1 AND "[120]8mm挡停缩回";
   IF #_w2 THEN "二站数据".电机正转 := TRUE; END_IF;
   IF #_w2 AND "二站数据".电机正转 THEN "手动模式数据".手动灌注总步骤 := 3.0; END_IF;
END_REGION
END_FUNCTION

FUNCTION "手动10mm流程" : Void   // FC7, LAD
{ S7_Optimized_Access := 'TRUE' }
VERSION : 0.1
   VAR_TEMP   // added for the SCL form of the ladder/FBD networks
      _w1 : Bool;
      _w2 : Bool;
   END_VAR
BEGIN

REGION Network 1
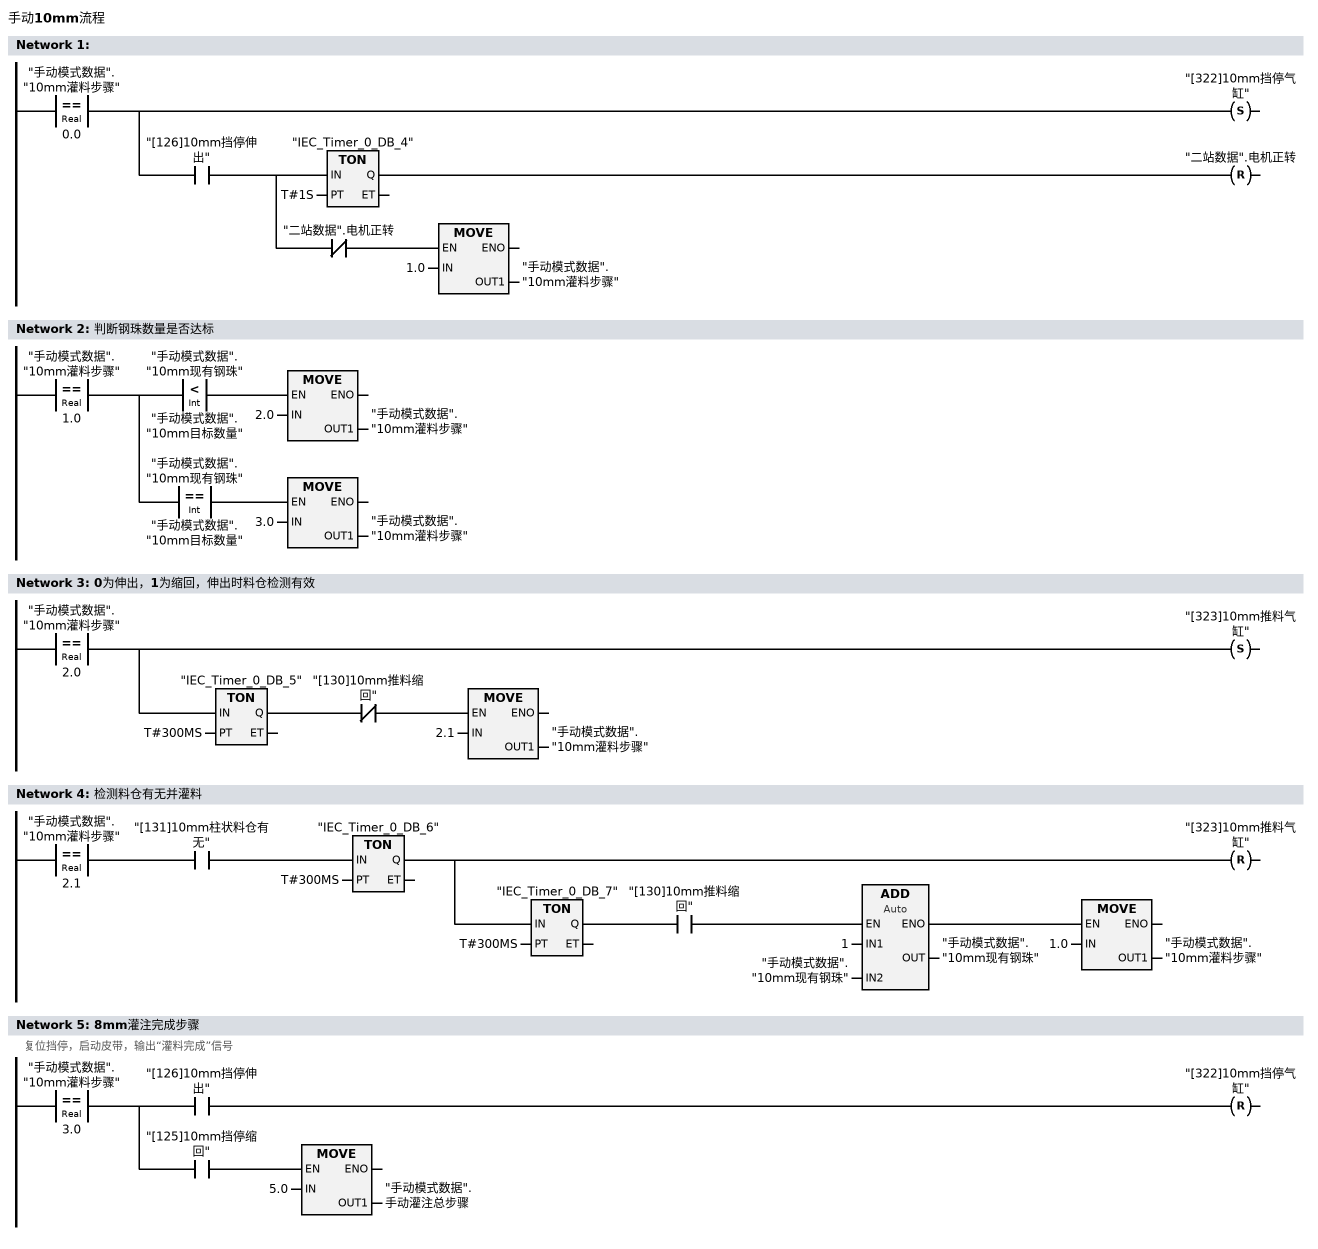
   #_w1 := "手动模式数据"."10mm灌料步骤" = 0.0;
   IF #_w1 THEN "[322]10mm挡停气缸" := TRUE; END_IF;
   #_w2 := #_w1 AND "[126]10mm挡停伸出";
   "IEC_Timer_0_DB_4".TON(IN := #_w2, PT := T#1S);
   IF "IEC_Timer_0_DB_4".Q THEN "二站数据".电机正转 := FALSE; END_IF;
   IF #_w2 AND NOT "二站数据".电机正转 THEN "手动模式数据"."10mm灌料步骤" := 1.0; END_IF;
END_REGION

REGION Network 2: 判断钢珠数量是否达标
   RUNG wire#powerrail
      { S7_Templates := "SrcType := Real" } EQ_Contact(in1 := "手动模式数据"."10mm灌料步骤", in2 := 1.0)
      wire#w1
      { S7_Templates := "SrcType := Int" } LT_Contact(in1 := "手动模式数据"."10mm现有钢珠", in2 := "手动模式数据"."10mm目标数量")
      Move(in := 2.0, out1 => "手动模式数据"."10mm灌料步骤")
   END_RUNG
   RUNG wire#w1
      { S7_Templates := "SrcType := Int" } EQ_Contact(in1 := "手动模式数据"."10mm现有钢珠", in2 := "手动模式数据"."10mm目标数量")
      Move(in := 3.0, out1 => "手动模式数据"."10mm灌料步骤")
   END_RUNG
   // the same network as SCL:
   #_w1 := "手动模式数据"."10mm灌料步骤" = 1.0;
   IF #_w1 AND ("手动模式数据"."10mm现有钢珠" < "手动模式数据"."10mm目标数量") THEN "手动模式数据"."10mm灌料步骤" := 2.0; END_IF;
   IF #_w1 AND ("手动模式数据"."10mm现有钢珠" = "手动模式数据"."10mm目标数量") THEN "手动模式数据"."10mm灌料步骤" := 3.0; END_IF;
END_REGION

REGION Network 3: 0为伸出，1为缩回，伸出时料仓检测有效
   #_w1 := "手动模式数据"."10mm灌料步骤" = 2.0;
   IF #_w1 THEN "[323]10mm推料气缸" := TRUE; END_IF;
   "IEC_Timer_0_DB_5".TON(IN := #_w1, PT := T#300MS);
   IF "IEC_Timer_0_DB_5".Q AND NOT "[130]10mm推料缩回" THEN "手动模式数据"."10mm灌料步骤" := 2.1; END_IF;
END_REGION

REGION Network 4: 检测料仓有无并灌料
   "IEC_Timer_0_DB_6".TON(IN := ("手动模式数据"."10mm灌料步骤" = 2.1) AND "[131]10mm柱状料仓有无", PT := T#300MS);
   IF "IEC_Timer_0_DB_6".Q THEN "[323]10mm推料气缸" := FALSE; END_IF;
   "IEC_Timer_0_DB_7".TON(IN := "IEC_Timer_0_DB_6".Q, PT := T#300MS);
   IF "IEC_Timer_0_DB_7".Q AND "[130]10mm推料缩回" THEN
       "手动模式数据"."10mm现有钢珠" := 1 + "手动模式数据"."10mm现有钢珠";
       "手动模式数据"."10mm灌料步骤" := 1.0;
   END_IF;
END_REGION

REGION Network 5: 8mm灌注完成步骤
   // 复位挡停，启动皮带，输出“灌料完成”信号
   RUNG wire#powerrail
      { S7_Templates := "SrcType := Real" } EQ_Contact(in1 := "手动模式数据"."10mm灌料步骤", in2 := 3.0)
      wire#w1
      Contact( "[126]10mm挡停伸出" )
      R_Coil( "[322]10mm挡停气缸" )
   END_RUNG
   RUNG wire#w1
      Contact( "[125]10mm挡停缩回" )
      Move(in := 5.0, out1 => "手动模式数据".手动灌注总步骤)
   END_RUNG
   // the same network as SCL:
   #_w1 := "手动模式数据"."10mm灌料步骤" = 3.0;
   IF #_w1 AND "[126]10mm挡停伸出" THEN "[322]10mm挡停气缸" := FALSE; END_IF;
   IF #_w1 AND "[125]10mm挡停缩回" THEN "手动模式数据".手动灌注总步骤 := 5.0; END_IF;
END_REGION
END_FUNCTION

// folder: 自动模式

FUNCTION "10mm流程" : Void   // FC5, LAD
{ S7_Optimized_Access := 'TRUE' }
VERSION : 0.1
   VAR_TEMP   // added for the SCL form of the ladder/FBD networks
      _w1 : Bool;
      _w2 : Bool;
   END_VAR
BEGIN

REGION Network 1: 皮带停止，准备下料
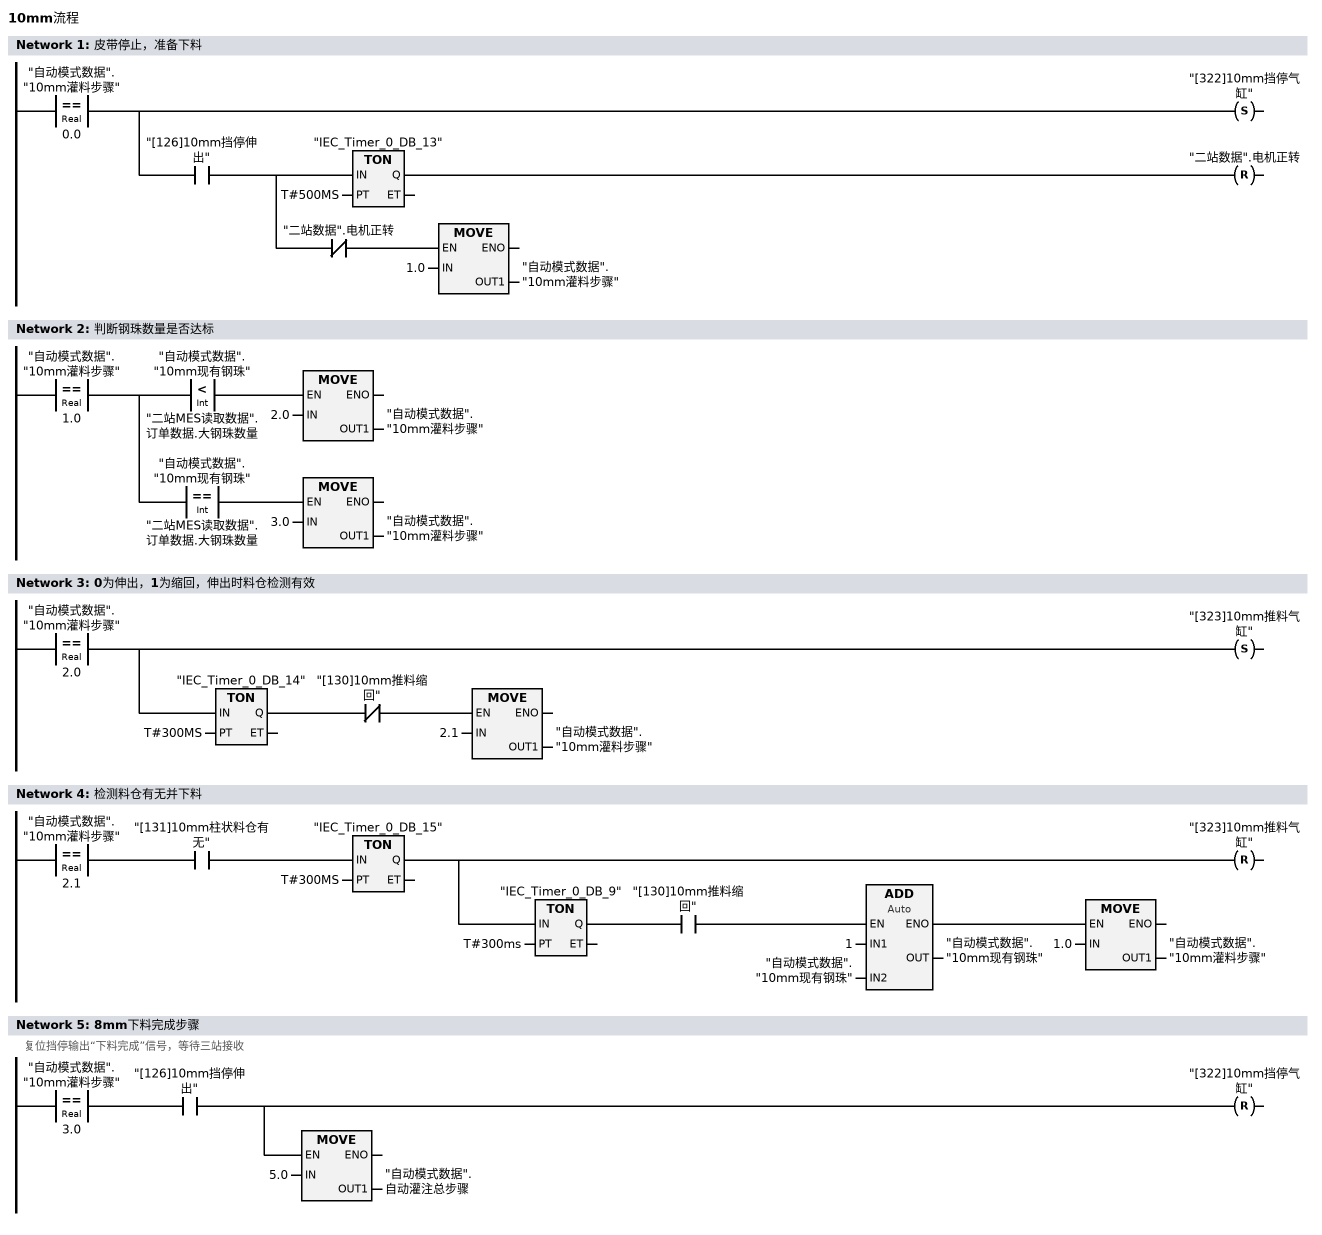
   #_w1 := "自动模式数据"."10mm灌料步骤" = 0.0;
   IF #_w1 THEN "[322]10mm挡停气缸" := TRUE; END_IF;
   #_w2 := #_w1 AND "[126]10mm挡停伸出";
   "IEC_Timer_0_DB_13".TON(IN := #_w2, PT := T#500MS);
   IF "IEC_Timer_0_DB_13".Q THEN "二站数据".电机正转 := FALSE; END_IF;
   IF #_w2 AND NOT "二站数据".电机正转 THEN "自动模式数据"."10mm灌料步骤" := 1.0; END_IF;
END_REGION

REGION Network 2: 判断钢珠数量是否达标
   RUNG wire#powerrail
      { S7_Templates := "SrcType := Real" } EQ_Contact(in1 := "自动模式数据"."10mm灌料步骤", in2 := 1.0)
      wire#w1
      { S7_Templates := "SrcType := Int" } LT_Contact(in1 := "自动模式数据"."10mm现有钢珠", in2 := "二站MES读取数据".订单数据.大钢珠数量)
      Move(in := 2.0, out1 => "自动模式数据"."10mm灌料步骤")
   END_RUNG
   RUNG wire#w1
      { S7_Templates := "SrcType := Int" } EQ_Contact(in1 := "自动模式数据"."10mm现有钢珠", in2 := "二站MES读取数据".订单数据.大钢珠数量)
      Move(in := 3.0, out1 => "自动模式数据"."10mm灌料步骤")
   END_RUNG
   // the same network as SCL:
   #_w1 := "自动模式数据"."10mm灌料步骤" = 1.0;
   IF #_w1 AND ("自动模式数据"."10mm现有钢珠" < "二站MES读取数据".订单数据.大钢珠数量) THEN "自动模式数据"."10mm灌料步骤" := 2.0; END_IF;
   IF #_w1 AND ("自动模式数据"."10mm现有钢珠" = "二站MES读取数据".订单数据.大钢珠数量) THEN "自动模式数据"."10mm灌料步骤" := 3.0; END_IF;
END_REGION

REGION Network 3: 0为伸出，1为缩回，伸出时料仓检测有效
   #_w1 := "自动模式数据"."10mm灌料步骤" = 2.0;
   IF #_w1 THEN "[323]10mm推料气缸" := TRUE; END_IF;
   "IEC_Timer_0_DB_14".TON(IN := #_w1, PT := T#300MS);
   IF "IEC_Timer_0_DB_14".Q AND NOT "[130]10mm推料缩回" THEN "自动模式数据"."10mm灌料步骤" := 2.1; END_IF;
END_REGION

REGION Network 4: 检测料仓有无并下料
   "IEC_Timer_0_DB_15".TON(IN := ("自动模式数据"."10mm灌料步骤" = 2.1) AND "[131]10mm柱状料仓有无", PT := T#300MS);
   IF "IEC_Timer_0_DB_15".Q THEN "[323]10mm推料气缸" := FALSE; END_IF;
   "IEC_Timer_0_DB_9".TON(IN := "IEC_Timer_0_DB_15".Q, PT := T#300ms);
   IF "IEC_Timer_0_DB_9".Q AND "[130]10mm推料缩回" THEN
       "自动模式数据"."10mm现有钢珠" := 1 + "自动模式数据"."10mm现有钢珠";
       "自动模式数据"."10mm灌料步骤" := 1.0;
   END_IF;
END_REGION

REGION Network 5: 8mm下料完成步骤
   // 复位挡停输出“下料完成”信号，等待三站接收
   RUNG wire#powerrail
      { S7_Templates := "SrcType := Real" } EQ_Contact(in1 := "自动模式数据"."10mm灌料步骤", in2 := 3.0)
      Contact( "[126]10mm挡停伸出" )
      wire#w1
      R_Coil( "[322]10mm挡停气缸" )
   END_RUNG
   RUNG wire#w1
      Move(in := 5.0, out1 => "自动模式数据".自动灌注总步骤)
   END_RUNG
   // the same network as SCL:
   #_w1 := ("自动模式数据"."10mm灌料步骤" = 3.0) AND "[126]10mm挡停伸出";
   IF #_w1 THEN
       "[322]10mm挡停气缸" := FALSE;
       "自动模式数据".自动灌注总步骤 := 5.0;
   END_IF;
END_REGION
END_FUNCTION

FUNCTION "8mm流程" : Void   // FC6, LAD
{ S7_Optimized_Access := 'TRUE' }
VERSION : 0.1
   VAR_TEMP   // added for the SCL form of the ladder/FBD networks
      _w1 : Bool;
      _w2 : Bool;
   END_VAR
BEGIN

REGION Network 1
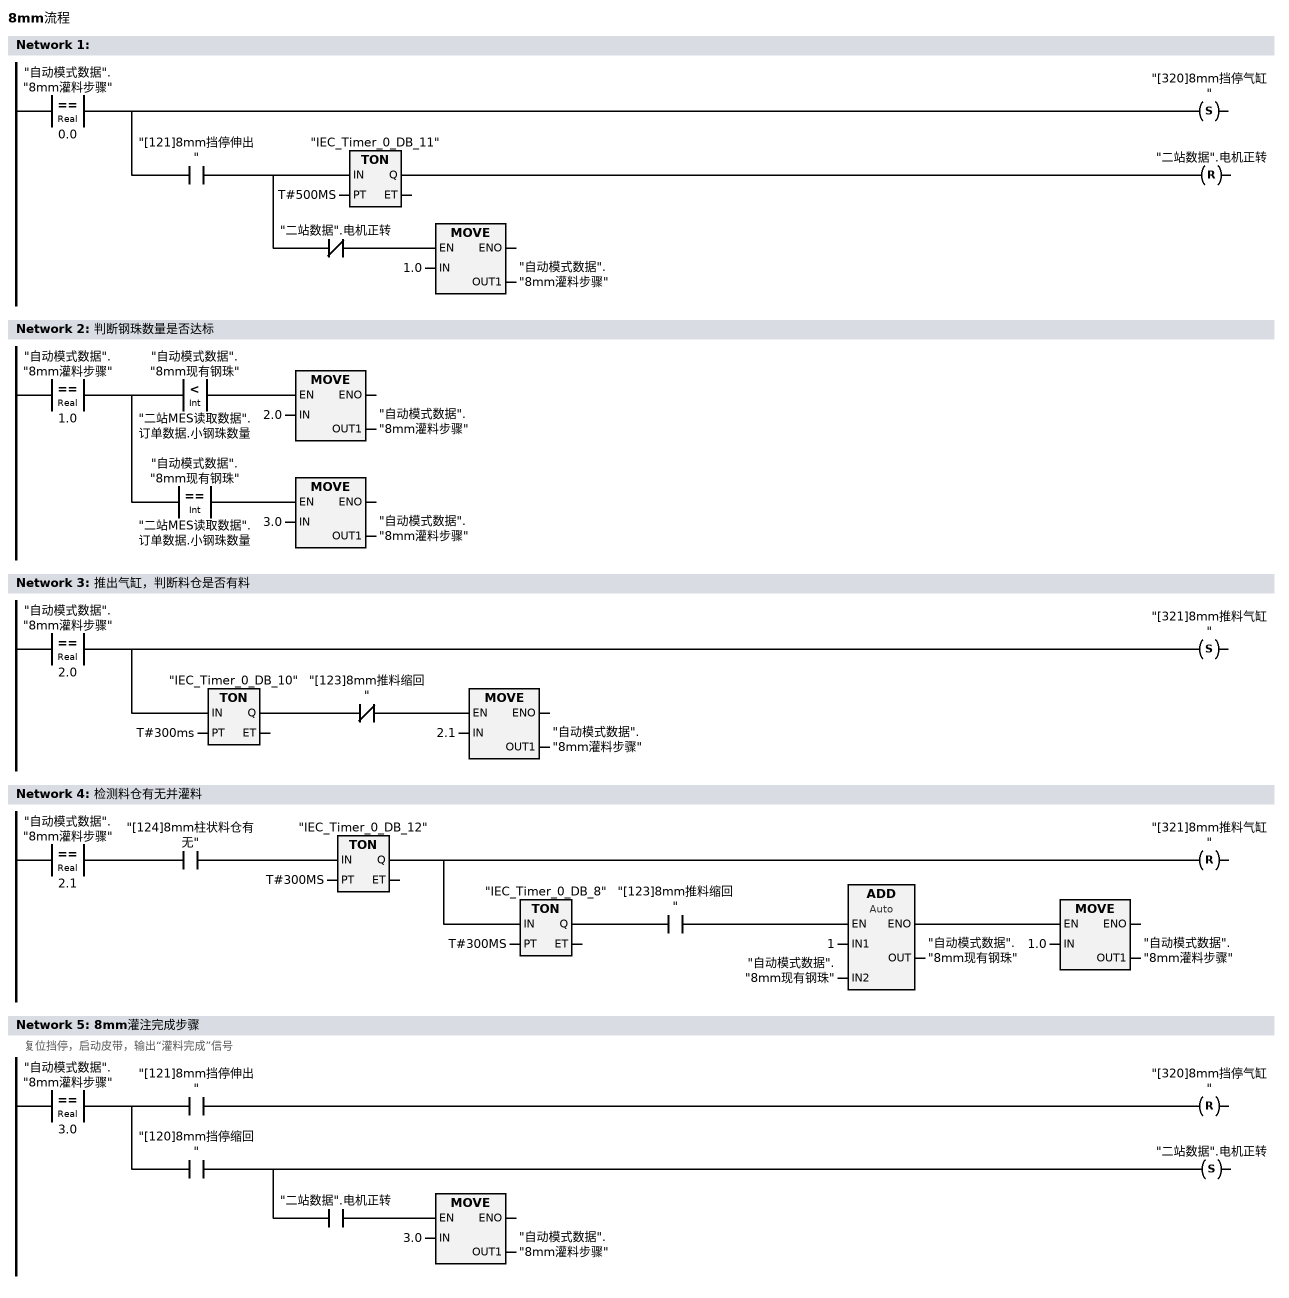
   #_w1 := "自动模式数据"."8mm灌料步骤" = 0.0;
   IF #_w1 THEN "[320]8mm挡停气缸" := TRUE; END_IF;
   #_w2 := #_w1 AND "[121]8mm挡停伸出";
   "IEC_Timer_0_DB_11".TON(IN := #_w2, PT := T#500MS);
   IF "IEC_Timer_0_DB_11".Q THEN "二站数据".电机正转 := FALSE; END_IF;
   IF #_w2 AND NOT "二站数据".电机正转 THEN "自动模式数据"."8mm灌料步骤" := 1.0; END_IF;
END_REGION

REGION Network 2: 判断钢珠数量是否达标
   RUNG wire#powerrail
      { S7_Templates := "SrcType := Real" } EQ_Contact(in1 := "自动模式数据"."8mm灌料步骤", in2 := 1.0)
      wire#w1
      { S7_Templates := "SrcType := Int" } LT_Contact(in1 := "自动模式数据"."8mm现有钢珠", in2 := "二站MES读取数据".订单数据.小钢珠数量)
      Move(in := 2.0, out1 => "自动模式数据"."8mm灌料步骤")
   END_RUNG
   RUNG wire#w1
      { S7_Templates := "SrcType := Int" } EQ_Contact(in1 := "自动模式数据"."8mm现有钢珠", in2 := "二站MES读取数据".订单数据.小钢珠数量)
      Move(in := 3.0, out1 => "自动模式数据"."8mm灌料步骤")
   END_RUNG
   // the same network as SCL:
   #_w1 := "自动模式数据"."8mm灌料步骤" = 1.0;
   IF #_w1 AND ("自动模式数据"."8mm现有钢珠" < "二站MES读取数据".订单数据.小钢珠数量) THEN "自动模式数据"."8mm灌料步骤" := 2.0; END_IF;
   IF #_w1 AND ("自动模式数据"."8mm现有钢珠" = "二站MES读取数据".订单数据.小钢珠数量) THEN "自动模式数据"."8mm灌料步骤" := 3.0; END_IF;
END_REGION

REGION Network 3: 推出气缸，判断料仓是否有料
   #_w1 := "自动模式数据"."8mm灌料步骤" = 2.0;
   IF #_w1 THEN "[321]8mm推料气缸" := TRUE; END_IF;
   "IEC_Timer_0_DB_10".TON(IN := #_w1, PT := T#300ms);
   IF "IEC_Timer_0_DB_10".Q AND NOT "[123]8mm推料缩回" THEN "自动模式数据"."8mm灌料步骤" := 2.1; END_IF;
END_REGION

REGION Network 4: 检测料仓有无并灌料
   "IEC_Timer_0_DB_12".TON(IN := ("自动模式数据"."8mm灌料步骤" = 2.1) AND "[124]8mm柱状料仓有无", PT := T#300MS);
   IF "IEC_Timer_0_DB_12".Q THEN "[321]8mm推料气缸" := FALSE; END_IF;
   "IEC_Timer_0_DB_8".TON(IN := "IEC_Timer_0_DB_12".Q, PT := T#300MS);
   IF "IEC_Timer_0_DB_8".Q AND "[123]8mm推料缩回" THEN
       "自动模式数据"."8mm现有钢珠" := 1 + "自动模式数据"."8mm现有钢珠";
       "自动模式数据"."8mm灌料步骤" := 1.0;
   END_IF;
END_REGION

REGION Network 5: 8mm灌注完成步骤
   // 复位挡停，启动皮带，输出“灌料完成”信号
   RUNG wire#powerrail
      { S7_Templates := "SrcType := Real" } EQ_Contact(in1 := "自动模式数据"."8mm灌料步骤", in2 := 3.0)
      wire#w1
      Contact( "[121]8mm挡停伸出" )
      R_Coil( "[320]8mm挡停气缸" )
   END_RUNG
   RUNG wire#w1
      Contact( "[120]8mm挡停缩回" )
      wire#w2
      S_Coil( "二站数据".电机正转 )
   END_RUNG
   RUNG wire#w2
      Contact( "二站数据".电机正转 )
      Move(in := 3.0, out1 => "自动模式数据"."8mm灌料步骤")
   END_RUNG
   // the same network as SCL:
   #_w1 := "自动模式数据"."8mm灌料步骤" = 3.0;
   IF #_w1 AND "[121]8mm挡停伸出" THEN "[320]8mm挡停气缸" := FALSE; END_IF;
   #_w2 := #_w1 AND "[120]8mm挡停缩回";
   IF #_w2 THEN "二站数据".电机正转 := TRUE; END_IF;
   IF #_w2 AND "二站数据".电机正转 THEN "自动模式数据"."8mm灌料步骤" := 3.0; END_IF;
END_REGION
END_FUNCTION

FUNCTION "自动下料流程" : Void   // FC10, LAD
{ S7_Optimized_Access := 'TRUE' }
VERSION : 0.1
   VAR_TEMP   // added for the SCL form of the ladder/FBD networks
      _w1 : Bool;
      _w2 : Bool;
   END_VAR
BEGIN

REGION Network 1: 复位
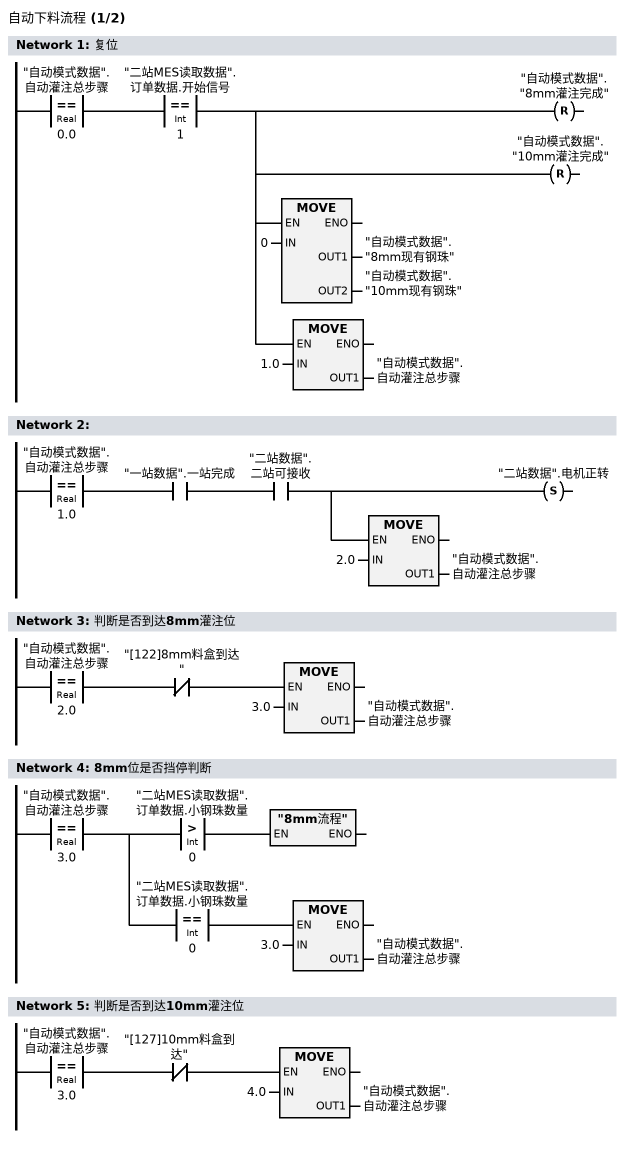
   RUNG wire#powerrail
      { S7_Templates := "SrcType := Real" } EQ_Contact(in1 := "自动模式数据".自动灌注总步骤, in2 := 0.0)
      { S7_Templates := "SrcType := Int" } EQ_Contact(in1 := "二站MES读取数据".订单数据.开始信号, in2 := 1)
      wire#w1
      R_Coil( "自动模式数据"."8mm灌注完成" )
   END_RUNG
   RUNG wire#w1
      R_Coil( "自动模式数据"."10mm灌注完成" )
   END_RUNG
   RUNG wire#w1
      Move(in := 0, out1 => "自动模式数据"."8mm现有钢珠", out2 => "自动模式数据"."10mm现有钢珠")
   END_RUNG
   RUNG wire#w1
      Move(in := 1.0, out1 => "自动模式数据".自动灌注总步骤)
   END_RUNG
   // the same network as SCL:
   IF ("自动模式数据".自动灌注总步骤 = 0.0) AND ("二站MES读取数据".订单数据.开始信号 = 1) THEN
       "自动模式数据"."8mm灌注完成" := FALSE;
       "自动模式数据"."10mm灌注完成" := FALSE;
       "自动模式数据"."8mm现有钢珠" := 0;
       "自动模式数据"."10mm现有钢珠" := 0;
       "自动模式数据".自动灌注总步骤 := 1.0;
   END_IF;
END_REGION

REGION Network 2
   RUNG wire#powerrail
      { S7_Templates := "SrcType := Real" } EQ_Contact(in1 := "自动模式数据".自动灌注总步骤, in2 := 1.0)
      Contact( "一站数据".一站完成 )
      Contact( "二站数据".二站可接收 )
      wire#w1
      S_Coil( "二站数据".电机正转 )
   END_RUNG
   RUNG wire#w1
      Move(in := 2.0, out1 => "自动模式数据".自动灌注总步骤)
   END_RUNG
   // the same network as SCL:
   IF ("自动模式数据".自动灌注总步骤 = 1.0) AND "一站数据".一站完成 AND "二站数据".二站可接收 THEN
       "二站数据".电机正转 := TRUE;
       "自动模式数据".自动灌注总步骤 := 2.0;
   END_IF;
END_REGION

REGION Network 3: 判断是否到达8mm灌注位
   RUNG wire#powerrail
      { S7_Templates := "SrcType := Real" } EQ_Contact(in1 := "自动模式数据".自动灌注总步骤, in2 := 2.0)
      I_Contact( "[122]8mm料盒到达" )
      Move(in := 3.0, out1 => "自动模式数据".自动灌注总步骤)
   END_RUNG
   // the same network as SCL:
   IF ("自动模式数据".自动灌注总步骤 = 2.0) AND NOT "[122]8mm料盒到达" THEN "自动模式数据".自动灌注总步骤 := 3.0; END_IF;
END_REGION

REGION Network 4: 8mm位是否挡停判断
   RUNG wire#powerrail
      { S7_Templates := "SrcType := Real" } EQ_Contact(in1 := "自动模式数据".自动灌注总步骤, in2 := 3.0)
      wire#w1
      { S7_Templates := "SrcType := Int" } GT_Contact(in1 := "二站MES读取数据".订单数据.小钢珠数量, in2 := 0)
      "8mm流程"()
   END_RUNG
   RUNG wire#w1
      { S7_Templates := "SrcType := Int" } EQ_Contact(in1 := "二站MES读取数据".订单数据.小钢珠数量, in2 := 0)
      Move(in := 3.0, out1 => "自动模式数据".自动灌注总步骤)
   END_RUNG
   // the same network as SCL:
   #_w1 := "自动模式数据".自动灌注总步骤 = 3.0;
   IF #_w1 AND ("二站MES读取数据".订单数据.小钢珠数量 > 0) THEN "8mm流程"(); END_IF;
   IF #_w1 AND ("二站MES读取数据".订单数据.小钢珠数量 = 0) THEN "自动模式数据".自动灌注总步骤 := 3.0; END_IF;
END_REGION

REGION Network 5: 判断是否到达10mm灌注位
   RUNG wire#powerrail
      { S7_Templates := "SrcType := Real" } EQ_Contact(in1 := "自动模式数据".自动灌注总步骤, in2 := 3.0)
      I_Contact( "[127]10mm料盒到达" )
      Move(in := 4.0, out1 => "自动模式数据".自动灌注总步骤)
   END_RUNG
   // the same network as SCL:
   IF ("自动模式数据".自动灌注总步骤 = 3.0) AND NOT "[127]10mm料盒到达" THEN "自动模式数据".自动灌注总步骤 := 4.0; END_IF;
END_REGION

REGION Network 6: 10mm位是否挡停判断
   // 10mm完成后只会复位挡停
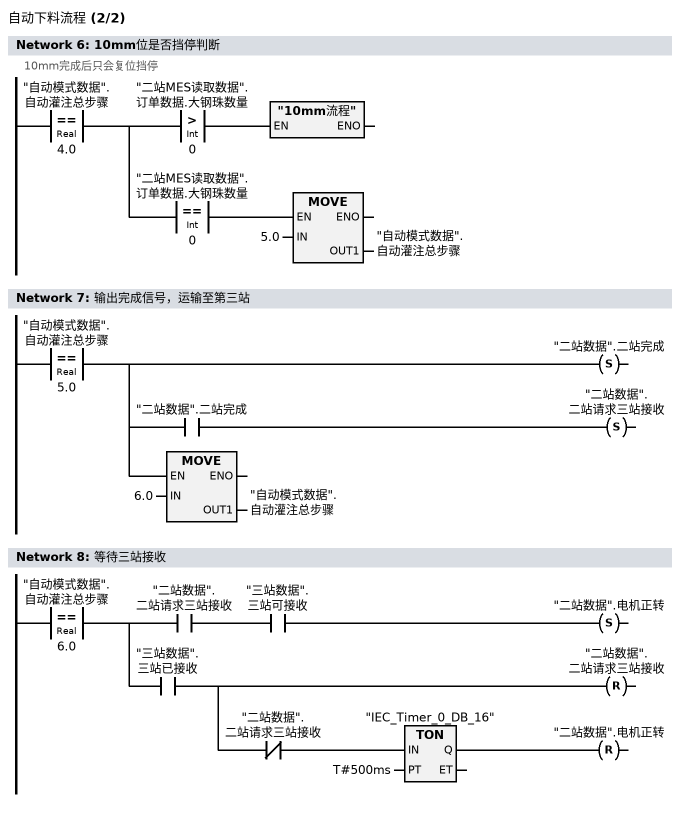
   RUNG wire#powerrail
      { S7_Templates := "SrcType := Real" } EQ_Contact(in1 := "自动模式数据".自动灌注总步骤, in2 := 4.0)
      wire#w1
      { S7_Templates := "SrcType := Int" } GT_Contact(in1 := "二站MES读取数据".订单数据.大钢珠数量, in2 := 0)
      "10mm流程"()
   END_RUNG
   RUNG wire#w1
      { S7_Templates := "SrcType := Int" } EQ_Contact(in1 := "二站MES读取数据".订单数据.大钢珠数量, in2 := 0)
      Move(in := 5.0, out1 => "自动模式数据".自动灌注总步骤)
   END_RUNG
   // the same network as SCL:
   #_w1 := "自动模式数据".自动灌注总步骤 = 4.0;
   IF #_w1 AND ("二站MES读取数据".订单数据.大钢珠数量 > 0) THEN "10mm流程"(); END_IF;
   IF #_w1 AND ("二站MES读取数据".订单数据.大钢珠数量 = 0) THEN "自动模式数据".自动灌注总步骤 := 5.0; END_IF;
END_REGION

REGION Network 7: 输出完成信号，运输至第三站
   RUNG wire#powerrail
      { S7_Templates := "SrcType := Real" } EQ_Contact(in1 := "自动模式数据".自动灌注总步骤, in2 := 5.0)
      wire#w1
      S_Coil( "二站数据".二站完成 )
   END_RUNG
   RUNG wire#w1
      Contact( "二站数据".二站完成 )
      S_Coil( "二站数据".二站请求三站接收 )
   END_RUNG
   RUNG wire#w1
      Move(in := 6.0, out1 => "自动模式数据".自动灌注总步骤)
   END_RUNG
   // the same network as SCL:
   #_w1 := "自动模式数据".自动灌注总步骤 = 5.0;
   IF #_w1 THEN "二站数据".二站完成 := TRUE; END_IF;
   IF #_w1 AND "二站数据".二站完成 THEN "二站数据".二站请求三站接收 := TRUE; END_IF;
   IF #_w1 THEN "自动模式数据".自动灌注总步骤 := 6.0; END_IF;
END_REGION

REGION Network 8: 等待三站接收
   #_w1 := "自动模式数据".自动灌注总步骤 = 6.0;
   IF #_w1 AND "二站数据".二站请求三站接收 AND "三站数据".三站可接收 THEN "二站数据".电机正转 := TRUE; END_IF;
   #_w2 := #_w1 AND "三站数据".三站已接收;
   IF #_w2 THEN "二站数据".二站请求三站接收 := FALSE; END_IF;
   "IEC_Timer_0_DB_16".TON(IN := #_w2 AND NOT "二站数据".二站请求三站接收, PT := T#500ms);
   IF "IEC_Timer_0_DB_16".Q THEN "二站数据".电机正转 := FALSE; END_IF;
END_REGION
END_FUNCTION

FUNCTION "数据转换以及检测" : Void   // FC14, LAD
{ S7_Optimized_Access := 'TRUE' }
VERSION : 0.1
BEGIN
END_FUNCTION

// folder: 通讯数据

FUNCTION "产线通讯" : Void   // FC2, LAD
{ S7_Optimized_Access := 'TRUE' }
VERSION : 0.1
BEGIN

REGION Network 1: 心跳
